// TwinCAT 3 PLC project BendingMachine
// ProgramVersion: 3.1.4026.27
// libraries:
//   Tc2_MC2, * (Beckhoff Automation GmbH)
//   Tc2_MC2_Drive, * (Beckhoff Automation GmbH)
//   Tc2_NCI, * (Beckhoff Automation GmbH)
//   Tc2_PlcInterpolation, * (Beckhoff Automation GmbH)
//   Tc2_Standard, * (Beckhoff Automation GmbH)
//   Tc2_SUPS, * (Beckhoff Automation GmbH)
//   Tc2_System, * (Beckhoff Automation GmbH)
//   Tc2_Utilities, * (Beckhoff Automation GmbH)
//   Tc3_JsonXml, * (Beckhoff Automation GmbH)
//   Tc3_MC2_AdvancedHoming, * (Beckhoff Automation GmbH)
// project tree:
//   DUTs/ ACTION_ENUM.TcDUT, AXIS_ENUM.TcDUT, CENTERING_ENUM.TcDUT, E_Alarm.TcDUT, EJECT_ENUM.TcDUT, OUTPUT_ACTION_ENUM.TcDUT, OUTPUT_ENUM.TcDUT, PRGSTATE_ENUM.TcDUT, ST_MpgEncoder.TcDUT, ST_TwoHandControl.TcDUT, TYPE_ACTION.TcDUT, TYPE_MACHINE_RX.TcDUT, TYPE_MACHINE_TX.TcDUT, TYPE_MACRO.TcDUT, TYPE_PARAMETERS.TcDUT, TYPE_POSITION.TcDUT, TYPE_SEQUENCE.TcDUT, TYPE_TASK.TcDUT
//   GVLs/ Alarms.TcGVL, Calibration.TcGVL, IO.TcGVL, Machine.TcGVL, ProgramDB.TcGVL, Safety.TcGVL, Size.TcGVL, Diag.TcGVL, Hmi.TcGVL
//   / PlcTask.TcTTO
//   POUs/ Clock.TcPOU, MAIN.TcPOU
//   Core/Valves/ SetMacro.TcPOU, WaitMacro.TcPOU, ST_Valve.TcDUT, ST_Input.TcDUT
//   POUs/Messages/ ClearAlarms.TcPOU, RaiseAlarm.TcPOU
//   POUs/MPG/ MPG_ReadStatus.TcPOU
//   Core/Nc/ FB_BuildGroups.TcPOU, FB_ClearInterpolationGroup.TcPOU, ST_AxisCfg.TcDUT, E_SeqCmd.TcDUT, E_SeqStep.TcDUT, FB_FeedTableBuilder.TcPOU, FB_SequenceRunner.TcPOU, E_NcChannelCmd.TcDUT, FB_NcChannels.TcPOU
//   POUs/TwoHand/ TwoHand_ReadStatus.TcPOU
//   Core/ Core_Param.TcGVL
//   Core/Cycle/ E_CycleState.TcDUT
//   Core/Diag/ E_CycleEndReason.TcDUT, ST_DiagEvent.TcDUT, ST_ChannelDiag.TcDUT, ST_Diag.TcDUT, FB_DiagLog.TcPOU
//   Core/Sync/ E_MFuncKind.TcDUT, E_MFuncOnError.TcDUT, ST_MFuncDef.TcDUT, F_MValve.TcPOU, F_MValveDirect.TcPOU, F_MSync.TcPOU, F_MSimple.TcPOU, FB_MFuncDispatcher.TcPOU
//   Machine/ E_Valve.TcDUT, Mach.TcGVL, FB_MachineConfig.TcPOU, FB_Centering.TcPOU, E_CenteringStep.TcDUT
//   Core/Axes/ FB_AxisModule.TcPOU, E_AxisAlarm.TcDUT
//   Core/Hmi/ E_HmiCommand.TcDUT, E_HmiResult.TcDUT, ST_HmiCmd.TcDUT, ST_HmiLive.TcDUT, ST_HmiAxisParam.TcDUT, ST_HmiParam.TcDUT, ST_HmiNamedItem.TcDUT, ST_HmiCfg.TcDUT, ST_HmiAxisSts.TcDUT, ST_HmiValveSts.TcDUT, ST_HmiSts.TcDUT, FB_HmiCommandHandler.TcPOU, FB_HmiWatchdog.TcPOU
// real-time tasks:
//   TASK PlcTask: cycle T#1ms, priority 20, ADS port 350
// motion (NC):
//   TASK NC-Task 1 SAF: cycle T#1ms, priority 1, ADS port 501
//   TASK NC-Task 1 SVB: cycle T#1ms, priority 8, ADS port 511
//   AXIS ERL (id 1)
//     General: UnitName=°
//     Dynamic: Acceleration=1780.713, Deceleration=1780.713, Jerk=5342.139
//     Velo: RefSearch=11.87142, RefSync=11.87142, SlowManual=59.3571, FastManual=356.1426, Fast=1187.142, Maximum=1187.142
//     OtherSettings: AllowMotionCmdToSlave=true
//     encoder EncType=8
//       EncPara: ScaleFactorNumerator=360, ScaleFactorDenominator=23068672, MaxCount=#xffffffff, ReferenceSystem=1
//         SoftEndMinControl: Enable=true, Range=-180
//         SoftEndMaxControl: Enable=true, Range=180
//     drive DrvType=9
//       DrvPara: MaxCount=#xffffffff, DriveControlDWord=#x00030100
//         Analog: VeloReferenz=1305.8562, VeloScale=1.02400649589962, TorqueSetpointScale=10, ScaleFactorActTorque=0.1
//         TimeComp: TaskDelayCycles=1
//     controller CtrType=1
//       CtrPara: PriorControlFactor=1
//         PosDiffControl: Enable=false
//         Observer: BandWidth=20
//   AXIS USEL (id 2)
//     Dynamic: Acceleration=1456.0155, Deceleration=1456.0155, Jerk=4368.0465
//     Velo: RefSearch=9.70677, RefSync=9.70677, SlowManual=12.5, FastManual=75, Fast=970.677, Maximum=970.677
//     OtherSettings: AllowMotionCmdToSlave=true
//     encoder EncType=8
//       EncPara: ScaleFactorNumerator=160, ScaleFactorDenominator=15728640, Offset=281.208719889323, Inverse=true, MaxCount=#xffffffff, ReferenceSystem=1
//         SoftEndMinControl: Enable=true, Range=66
//         SoftEndMaxControl: Enable=true, Range=1725
//     drive DrvType=9
//       DrvPara: Inverse=true, MaxCount=#xffffffff, DriveControlDWord=#x00030100
//         Analog: VeloReferenz=1067.7447, VeloScale=1.02400649589962, TorqueSetpointScale=10, ScaleFactorActTorque=0.1
//         TimeComp: TaskDelayCycles=1
//     controller CtrType=1
//       CtrPara: PriorControlFactor=1
//         Observer: BandWidth=20
//   AXIS ERR (id 3)
//     General: UnitName=°
//     Dynamic: Acceleration=1780.713, Deceleration=1780.713, Jerk=5342.139
//     Velo: RefSearch=11.87142, RefSync=11.87142, SlowManual=59.3571, FastManual=356.1426, Fast=1187.142, Maximum=1187.142
//     OtherSettings: AllowMotionCmdToSlave=true
//     encoder EncType=8
//       EncPara: ScaleFactorNumerator=360, ScaleFactorDenominator=23068672, Offset=78.9122668179599, MaxCount=#xffffffff, ReferenceSystem=1
//         SoftEndMinControl: Enable=true, Range=-180
//         SoftEndMaxControl: Enable=true, Range=180
//     drive DrvType=9
//       DrvPara: MaxCount=#xffffffff, DriveControlDWord=#x00030100
//         Analog: VeloReferenz=1305.8562, VeloScale=1.02400649589962, TorqueSetpointScale=10, ScaleFactorActTorque=0.1
//         TimeComp: TaskDelayCycles=1
//     controller CtrType=1
//       CtrPara: PriorControlFactor=1
//         Observer: BandWidth=20
//   AXIS USER (id 4)
//     Dynamic: Acceleration=1456.0155, Deceleration=1456.0155, Jerk=4368.0465
//     Velo: RefSearch=9.70677, RefSync=9.70677, SlowManual=12.5, FastManual=75, Fast=970.677, Maximum=970.677
//     OtherSettings: AllowMotionCmdToSlave=true
//     encoder EncType=8
//       EncPara: ScaleFactorNumerator=160, ScaleFactorDenominator=15728640, Offset=543.740122477214, Inverse=true, MaxCount=#xffffffff, ReferenceSystem=1
//         SoftEndMinControl: Enable=true, Range=66
//         SoftEndMaxControl: Enable=true, Range=1725
//     drive DrvType=9
//       DrvPara: Inverse=true, MaxCount=#xffffffff, DriveControlDWord=#x00030100
//         Analog: VeloReferenz=1067.7447, VeloScale=1.02400649589962, TorqueSetpointScale=10, ScaleFactorActTorque=0.1
//         TimeComp: TaskDelayCycles=1
//     controller CtrType=1
//       CtrPara: PriorControlFactor=1
//         Observer: BandWidth=20
//   AXIS UR (id 5)
//     General: UnitName=°
//     Dynamic: Acceleration=546.441, Deceleration=546.441, Jerk=1639.323
//     Velo: RefSearch=3.64294, RefSync=3.64294, SlowManual=18.2147, FastManual=109.2882, Fast=364.294, Maximum=364.294
//     OtherSettings: AllowMotionCmdToSlave=true
//     encoder EncType=8
//       EncPara: ScaleFactorNumerator=360, ScaleFactorDenominator=57671680, Offset=-105.826067837802, MaxCount=#xffffffff, ReferenceSystem=1
//         SoftEndMinControl: Enable=true, Range=-95
//         SoftEndMaxControl: Enable=true, Range=95
//     drive DrvType=9
//       DrvPara: MaxCount=#xffffffff, DriveControlDWord=#x00030100
//         Analog: VeloReferenz=400.7234, VeloScale=1.02400649589962, TorqueSetpointScale=10, ScaleFactorActTorque=0.1
//         TimeComp: TaskDelayCycles=1
//     controller CtrType=1
//       CtrPara: PriorControlFactor=1
//         Observer: BandWidth=20
//   AXIS UR SIM (id 6)
//     OtherSettings: AllowMotionCmdToSlave=true
//     encoder EncType=1
//     drive DrvType=5
//       Analog: TorqueSetpointScale=10, ScaleFactorActTorque=0.1
//       TimeComp: TaskDelayCycles=1
//     controller CtrType=1
//       CtrPara: PriorControlFactor=1
//         Observer: BandWidth=20
// I/O:
//   DEVICE Device 1 (EtherCAT), AmsNetId 192.168.1.106.2.1
//     Term 21 (EK1100) [EK1100 EtherCAT Coupler (2A E-Bus)]
//       Term 22 (EL6070-0033) [EL6070-0033 1Ch. Licence key terminal, individual licences]
//       Term 23 (EL1409) [EL1409 16Ch. Dig. Input 24V, 3ms]
//       Term 24 (EL1409) [EL1409 16Ch. Dig. Input 24V, 3ms]
//       Term 25 (EL2409) [EL2409 16Ch. Dig. Output 24V, 0.5A]
//       Term 26 (EK1322) [EK1322 2-port EtherCAT P junction with feed-in]
//         Box 27 (EPP1809-0022) [EPP1809-0022 16 Ch. Dig. Input 24V, 3ms, M8]
//         Box 28 (EPP1809-0022) [EPP1809-0022 16 Ch. Dig. Input 24V, 3ms, M8]
//       Term 29 (EL9410) [EL9410 E-Bus Power Supplier  (Diagnostics)]
//       Term 30 (EL6910) [EL6910, TwinSAFE PLC]
//       Term 31 (EL1918) [EL1918, 8Ch. Safety Input 24V, TwinSAFE]
//         modules: Module 1 (FSOE), Module 2 (FSLOGIC)
//       Term 32 (EL1918) [EL1918, 8Ch. Safety Input 24V, TwinSAFE]
//         modules: Module 1 (FSOE), Module 2 (FSLOGIC)
//       Term 33 (EL2904) [EL2904, 4 Ch. Safety Output 24V, 0.5A, TwinSAFE]
//         modules: Module 1 (FSOES), Module 2 (DO)
//       Term 34 (EK1110) [EK1110 EtherCAT extension]
//     Drive 35 (AX5206-0000-0216) [AX5206-0000-0216 EtherCAT Drive (SoE, 2 Ch.)]
//       Term 36 (AX5805) [AX5805 (Safety Drive Option)]
//         modules: Module 1 (Safety Process Data, 2 axis), Module 2 (Standard Process Data, 2 axis)
//     Drive 37 (AX5206-0000-0216) [AX5206-0000-0216 EtherCAT Drive (SoE, 2 Ch.)]
//       Term 38 (AX5805) [AX5805 (Safety Drive Option)]
//         modules: Module 1 (Safety Process Data, 2 axis), Module 2 (Standard Process Data, 2 axis)
//     Box 41 (EX260-SEC1) [EX260-SEC1 EtherCAT SI Unit (32DO_PNP) Rev1.2]
//     Box 42 (EX260-SEC1) [EX260-SEC1 EtherCAT SI Unit (32DO_PNP) Rev1.2]
//     Drive 39 (AX5103-0000-0216) [AX5103-0000-0216 EtherCAT Drive (SoE, 1 Ch.)]
//       Term 40 (AX5805) [AX5805 (Safety Drive Option)]
//         modules: Module 1 (Safety Process Data, 1 axis), Module 2 (Standard Process Data, 1 axis)
// variable links:
//   Device 1 (EtherCAT) <-> Device 1 (EtherCAT)/Drive 35 (AX5206-0000-0216)/Term 36 (AX5805)
//     Term 21 (EK1100)/Term 30 (EL6910)/ConnectionInputs/Message_184 TxPDO <-> Module 1 (Safety Process Data, 2 axis)/Outputs (Controlword)/FSOE
//     Term 21 (EK1100)/Term 30 (EL6910)/ConnectionOutputs/Message_184 RxPDO <-> Module 1 (Safety Process Data, 2 axis)/Inputs (Statusword)/FSOE
//   Device 1 (EtherCAT) <-> Device 1 (EtherCAT)/Drive 37 (AX5206-0000-0216)/Term 38 (AX5805)
//     Term 21 (EK1100)/Term 30 (EL6910)/ConnectionInputs/Message_183 TxPDO <-> Module 1 (Safety Process Data, 2 axis)/Outputs (Controlword)/FSOE
//     Term 21 (EK1100)/Term 30 (EL6910)/ConnectionOutputs/Message_183 RxPDO <-> Module 1 (Safety Process Data, 2 axis)/Inputs (Statusword)/FSOE
//   Device 1 (EtherCAT) <-> Device 1 (EtherCAT)/Drive 39 (AX5103-0000-0216)/Term 40 (AX5805)
//     Term 21 (EK1100)/Term 30 (EL6910)/ConnectionInputs/Message_191 TxPDO <-> Module 1 (Safety Process Data, 1 axis)/Outputs (Controlword)/FSOE
//     Term 21 (EK1100)/Term 30 (EL6910)/ConnectionOutputs/Message_191 RxPDO <-> Module 1 (Safety Process Data, 1 axis)/Inputs (Statusword)/FSOE
//   Device 1 (EtherCAT) <-> Device 1 (EtherCAT)/Term 21 (EK1100)/Term 31 (EL1918)
//     Term 21 (EK1100)/Term 30 (EL6910)/ConnectionInputs/Message_195 TxPDO <-> Module 1 (FSOE)/FSoE Outputs/FSOE
//     Term 21 (EK1100)/Term 30 (EL6910)/ConnectionOutputs/Message_195 RxPDO <-> Module 1 (FSOE)/FSoE Inputs/FSOE
//   Device 1 (EtherCAT) <-> Device 1 (EtherCAT)/Term 21 (EK1100)/Term 32 (EL1918)
//     Term 21 (EK1100)/Term 30 (EL6910)/ConnectionInputs/Message_196 TxPDO <-> Module 1 (FSOE)/FSoE Outputs/FSOE
//     Term 21 (EK1100)/Term 30 (EL6910)/ConnectionOutputs/Message_196 RxPDO <-> Module 1 (FSOE)/FSoE Inputs/FSOE
//   Device 1 (EtherCAT) <-> Device 1 (EtherCAT)/Term 21 (EK1100)/Term 33 (EL2904)
//     Term 21 (EK1100)/Term 30 (EL6910)/ConnectionInputs/Message_197 TxPDO <-> Module 1 (FSOES)/RxPDO/FSOE
//     Term 21 (EK1100)/Term 30 (EL6910)/ConnectionOutputs/Message_197 RxPDO <-> Module 1 (FSOES)/TxPDO/FSOE
//   NC-Task 1 SAF/Axes/ERL <-> Device 1 (EtherCAT)/Drive 35 (AX5206-0000-0216)
//     Drive/Inputs/In/nDataIn1 <-> AT 1/Following distance
//     Drive/Inputs/In/nDataIn3[0] <-> AT 1/Torque/force feedback value
//     Drive/Inputs/In/nDcOutputTime <-> InfoData/DcOutputShift
//     Drive/Inputs/In/nState1 <-> AT 1/Drive status word @bit 8
//     Drive/Inputs/In/nState2 <-> AT 1/Drive status word
//     Drive/Inputs/In/nState4 @bit 1 <-> WcState/InputToggle
//     Drive/Inputs/In/nState4 <-> WcState/WcState
//     Drive/Outputs/Out/nCtrl1 <-> MDT 1/Master control word @bit 8
//     Drive/Outputs/Out/nDataOut1 <-> MDT 1/Position command value
//     Enc/Inputs/In/nDataIn1 <-> AT 1/Position feedback 1 value
//     Enc/Inputs/In/nDcInputTime <-> InfoData/DcInputShift
//     Enc/Inputs/In/nState4 @bit 1 <-> WcState/InputToggle
//     Enc/Inputs/In/nState4 <-> WcState/WcState
//   NC-Task 1 SAF/Axes/ERR <-> Device 1 (EtherCAT)/Drive 37 (AX5206-0000-0216)
//     Drive/Inputs/In/nDataIn1 <-> AT 1/Following distance
//     Drive/Inputs/In/nDataIn3[0] <-> AT 1/Torque/force feedback value
//     Drive/Inputs/In/nDcOutputTime <-> InfoData/DcOutputShift
//     Drive/Inputs/In/nState1 <-> AT 1/Drive status word @bit 8
//     Drive/Inputs/In/nState2 <-> AT 1/Drive status word
//     Drive/Inputs/In/nState4 @bit 1 <-> WcState/InputToggle
//     Drive/Inputs/In/nState4 <-> WcState/WcState
//     Drive/Outputs/Out/nCtrl1 <-> MDT 1/Master control word @bit 8
//     Drive/Outputs/Out/nDataOut1 <-> MDT 1/Position command value
//     Enc/Inputs/In/nDataIn1 <-> AT 1/Position feedback 1 value
//     Enc/Inputs/In/nDcInputTime <-> InfoData/DcInputShift
//     Enc/Inputs/In/nState4 @bit 1 <-> WcState/InputToggle
//     Enc/Inputs/In/nState4 <-> WcState/WcState
//   NC-Task 1 SAF/Axes/UR <-> Device 1 (EtherCAT)/Drive 39 (AX5103-0000-0216)
//     Drive/Inputs/In/nDataIn1 <-> AT/Following distance
//     Drive/Inputs/In/nDataIn3[0] <-> AT/Torque/force feedback value
//     Drive/Inputs/In/nDcOutputTime <-> InfoData/DcOutputShift
//     Drive/Inputs/In/nState1 <-> AT/Drive status word @bit 8
//     Drive/Inputs/In/nState2 <-> AT/Drive status word
//     Drive/Inputs/In/nState4 @bit 1 <-> WcState/InputToggle
//     Drive/Inputs/In/nState4 <-> WcState/WcState
//     Drive/Outputs/Out/nCtrl1 <-> MDT/Master control word @bit 8
//     Drive/Outputs/Out/nDataOut1 <-> MDT/Position command value
//     Enc/Inputs/In/nDataIn1 <-> AT/Position feedback 1 value
//     Enc/Inputs/In/nDcInputTime <-> InfoData/DcInputShift
//     Enc/Inputs/In/nState4 @bit 1 <-> WcState/InputToggle
//     Enc/Inputs/In/nState4 <-> WcState/WcState
//   NC-Task 1 SAF/Axes/USEL <-> Device 1 (EtherCAT)/Drive 35 (AX5206-0000-0216)
//     Drive/Inputs/In/nDataIn1 <-> AT 2/Following distance
//     Drive/Inputs/In/nDataIn3[0] <-> AT 2/Torque/force feedback value
//     Drive/Inputs/In/nDcOutputTime <-> InfoData/DcOutputShift
//     Drive/Inputs/In/nState1 <-> AT 2/Drive status word @bit 8
//     Drive/Inputs/In/nState2 <-> AT 2/Drive status word
//     Drive/Inputs/In/nState4 @bit 1 <-> WcState/InputToggle
//     Drive/Inputs/In/nState4 <-> WcState/WcState
//     Drive/Outputs/Out/nCtrl1 <-> MDT 2/Master control word @bit 8
//     Drive/Outputs/Out/nDataOut1 <-> MDT 2/Position command value
//     Enc/Inputs/In/nDataIn1 <-> AT 2/Position feedback 1 value
//     Enc/Inputs/In/nDcInputTime <-> InfoData/DcInputShift
//     Enc/Inputs/In/nState4 @bit 1 <-> WcState/InputToggle
//     Enc/Inputs/In/nState4 <-> WcState/WcState
//   NC-Task 1 SAF/Axes/USER <-> Device 1 (EtherCAT)/Drive 37 (AX5206-0000-0216)
//     Drive/Inputs/In/nDataIn1 <-> AT 2/Following distance
//     Drive/Inputs/In/nDataIn3[0] <-> AT 2/Torque/force feedback value
//     Drive/Inputs/In/nDcOutputTime <-> InfoData/DcOutputShift
//     Drive/Inputs/In/nState1 <-> AT 2/Drive status word @bit 8
//     Drive/Inputs/In/nState2 <-> AT 2/Drive status word
//     Drive/Inputs/In/nState4 @bit 1 <-> WcState/InputToggle
//     Drive/Inputs/In/nState4 <-> WcState/WcState
//     Drive/Outputs/Out/nCtrl1 <-> MDT 2/Master control word @bit 8
//     Drive/Outputs/Out/nDataOut1 <-> MDT 2/Position command value
//     Enc/Inputs/In/nDataIn1 <-> AT 2/Position feedback 1 value
//     Enc/Inputs/In/nDcInputTime <-> InfoData/DcInputShift
//     Enc/Inputs/In/nState4 @bit 1 <-> WcState/InputToggle
//     Enc/Inputs/In/nState4 <-> WcState/WcState
//   BendingMachine/BendingMachine Instance <-> Device 1 (EtherCAT)/Box 41 (EX260-SEC1)
//     PlcTask Outputs/IO.smc1[{0..3}] <-> Byte {0..3}/Output  (4 links)
//   BendingMachine/BendingMachine Instance <-> Device 1 (EtherCAT)/Box 42 (EX260-SEC1)
//     PlcTask Outputs/IO.smc2[{0..3}] <-> Byte {0..3}/Output  (4 links)
//   BendingMachine/BendingMachine Instance <-> Device 1 (EtherCAT)/Drive 35 (AX5206-0000-0216)
//     PlcTask Inputs/MAIN.stMpgEncoder.diRowPositionFeedBack <-> AT 1/Position feedback 2 value (external feedback)
//   BendingMachine/BendingMachine Instance <-> Device 1 (EtherCAT)/Term 21 (EK1100)/Term 23 (EL1409)
//     PlcTask Inputs/IO.clampIn <-> DIP Inputs/Input Channel 14
//     PlcTask Inputs/IO.clampOpen <-> DIP Inputs/Input Channel 13
//     PlcTask Inputs/IO.fixedClampEncode <-> DIP Inputs/Input Channel 15
//     PlcTask Inputs/IO.mobileClampEncode <-> DIP Inputs/Input Channel 16
//     PlcTask Inputs/MAIN.stMpgEncoder.diButton1 <-> DIP Inputs/Input Channel 1
//     PlcTask Inputs/MAIN.stMpgEncoder.diButton2 <-> DIP Inputs/Input Channel 2
//     PlcTask Inputs/MAIN.stMpgEncoder.diButton3 <-> DIP Inputs/Input Channel 3
//     PlcTask Inputs/MAIN.stMpgEncoder.diSelector1Bit1 <-> DIP Inputs/Input Channel 4
//     PlcTask Inputs/MAIN.stMpgEncoder.diSelector1Bit2 <-> DIP Inputs/Input Channel 5
//     PlcTask Inputs/MAIN.stMpgEncoder.diSelector1Bit3 <-> DIP Inputs/Input Channel 6
//     PlcTask Inputs/MAIN.stMpgEncoder.diSelector2Bit1 <-> DIP Inputs/Input Channel 7
//     PlcTask Inputs/MAIN.stMpgEncoder.diSelector2Bit2 <-> DIP Inputs/Input Channel 8
//     PlcTask Inputs/MAIN.stTwoHandControl.diStartButton <-> DIP Inputs/Input Channel 9
//     PlcTask Inputs/MAIN.stTwoHandControl.diStopButton <-> DIP Inputs/Input Channel 10
//     PlcTask Inputs/Safety.PulsanteResetBarriere <-> DIP Inputs/Input Channel 12
//     PlcTask Inputs/Safety.PulsanteResetEmergenza <-> DIP Inputs/Input Channel 11
//   BendingMachine/BendingMachine Instance <-> Device 1 (EtherCAT)/Term 21 (EK1100)/Term 24 (EL1409)
//     PlcTask Inputs/IO.cabinetThermostat <-> DIP Inputs/Input Channel 10
//     PlcTask Inputs/IO.chillerAlarm <-> DIP Inputs/Input Channel 5
//     PlcTask Inputs/IO.chillerMagnetTrip <-> DIP Inputs/Input Channel 6
//     PlcTask Inputs/IO.doorLeftClosed <-> DIP Inputs/Input Channel 7
//     PlcTask Inputs/IO.doorRightClosed <-> DIP Inputs/Input Channel 8
//     PlcTask Inputs/IO.fuseAlarm <-> DIP Inputs/Input Channel 1
//     PlcTask Inputs/IO.leftAxisMagnetTrip <-> DIP Inputs/Input Channel 2
//     PlcTask Inputs/IO.pressureSwMinPressure <-> DIP Inputs/Input Channel 9
//     PlcTask Inputs/IO.rightAxisMagnetTrip <-> DIP Inputs/Input Channel 3
//     PlcTask Inputs/IO.ur2MagnetTrip <-> DIP Inputs/Input Channel 4
//   BendingMachine/BendingMachine Instance <-> Device 1 (EtherCAT)/Term 21 (EK1100)/Term 25 (EL2409)
//     PlcTask Outputs/IO.chillerEnabled <-> Channel 10/Output
//     PlcTask Outputs/IO.fuseReset <-> Channel 9/Output
//     PlcTask Outputs/IO.spiaPulsanteStart <-> Channel 7/Output
//     PlcTask Outputs/IO.spiaPulsanteStop <-> Channel 8/Output
//     PlcTask Outputs/IO.turretGreen <-> Channel 2/Output
//     PlcTask Outputs/IO.turretRed <-> Channel 1/Output
//     PlcTask Outputs/IO.turretSiren <-> Channel 4/Output
//     PlcTask Outputs/IO.turretYellow <-> Channel 3/Output
//     PlcTask Outputs/Safety.SpiaPulsanteRipristinoBarriere <-> Channel 6/Output
//     PlcTask Outputs/Safety.SpiaPulsanteRipristinoSicurezze <-> Channel 5/Output
//   BendingMachine/BendingMachine Instance <-> Device 1 (EtherCAT)/Term 21 (EK1100)/Term 26 (EK1322)/Box 27 (EPP1809-0022)
//     PlcTask Inputs/IO.centering1LeftIn <-> Channel 10/Input
//     PlcTask Inputs/IO.centering2LeftIn <-> Channel 9/Input
//     PlcTask Inputs/IO.centering3LeftIn <-> Channel 12/Input
//     PlcTask Inputs/IO.centering4LeftIn <-> Channel 11/Input
//     PlcTask Inputs/IO.epLeftBendUp <-> Channel 6/Input
//     PlcTask Inputs/IO.epLeftIn <-> Channel 5/Input
//     PlcTask Inputs/IO.erLeftIn <-> Channel 4/Input
//     PlcTask Inputs/IO.erLeftOut <-> Channel 3/Input
//     PlcTask Inputs/IO.useLeftDown <-> Channel 2/Input
//     PlcTask Inputs/IO.useLeftUp <-> Channel 1/Input
//   BendingMachine/BendingMachine Instance <-> Device 1 (EtherCAT)/Term 21 (EK1100)/Term 26 (EK1322)/Box 28 (EPP1809-0022)
//     PlcTask Inputs/IO.epRightBendUp <-> Channel 6/Input
//     PlcTask Inputs/IO.epRightIn <-> Channel 5/Input
//     PlcTask Inputs/IO.erRightIn <-> Channel 4/Input
//     PlcTask Inputs/IO.erRightOut <-> Channel 3/Input
//     PlcTask Inputs/IO.useRightDown <-> Channel 2/Input
//     PlcTask Inputs/IO.useRighttUp <-> Channel 1/Input
//   BendingMachine/BendingMachine Instance <-> Device 1 (EtherCAT)/Term 21 (EK1100)/Term 30 (EL6910)
//     PlcTask Inputs/MAIN.stMpgEncoder.diSafetySwitch <-> StandardInputs/Standard Out Var 64
//     PlcTask Inputs/MAIN.stTwoHandControl.diSafetySwitch <-> StandardInputs/Standard Out Var 60
//     PlcTask Inputs/MAIN.stTwoHandControl.diTwoHand <-> StandardInputs/Standard Out Var 65
//     PlcTask Inputs/Safety.AbilitazionePeriferiche <-> StandardInputs/Standard Out Var 50
//     PlcTask Inputs/Safety.BarriereResettate <-> StandardInputs/Standard Out Var 62
//     PlcTask Inputs/Safety.ComErr <-> StandardInputs/Standard Out Var 13
//     PlcTask Inputs/Safety.ComStartup <-> StandardInputs/Standard Out Var 14
//     PlcTask Inputs/Safety.ERL_Error <-> StandardInputs/Standard Out Var 93
//     PlcTask Inputs/Safety.ERL_SDI_n <-> StandardInputs/Standard Out Var 92
//     PlcTask Inputs/Safety.ERL_SDI_p <-> StandardInputs/Standard Out Var 91
//     PlcTask Inputs/Safety.ERL_SOS <-> StandardInputs/Standard Out Var 89
//     PlcTask Inputs/Safety.ERL_SSM1 <-> StandardInputs/Standard Out Var 87
//     PlcTask Inputs/Safety.ERL_SSM2 <-> StandardInputs/Standard Out Var 88
//     PlcTask Inputs/Safety.ERL_SSR <-> StandardInputs/Standard Out Var 90
//     PlcTask Inputs/Safety.ERL_STO <-> StandardInputs/Standard Out Var 86
//     PlcTask Inputs/Safety.ERR_Error <-> StandardInputs/Standard Out Var 112
//     PlcTask Inputs/Safety.ERR_SDI_n <-> StandardInputs/Standard Out Var 113
//     PlcTask Inputs/Safety.ERR_SDI_p <-> StandardInputs/Standard Out Var 103
//     PlcTask Inputs/Safety.ERR_SOS <-> StandardInputs/Standard Out Var 104
//     PlcTask Inputs/Safety.ERR_SSM1 <-> StandardInputs/Standard Out Var 105
//     PlcTask Inputs/Safety.ERR_SSM2 <-> StandardInputs/Standard Out Var 106
//     PlcTask Inputs/Safety.ERR_SSR <-> StandardInputs/Standard Out Var 107
//     PlcTask Inputs/Safety.ERR_SSR2 <-> StandardInputs/Standard Out Var 182
//     PlcTask Inputs/Safety.ERR_STO <-> StandardInputs/Standard Out Var 108
//     PlcTask Inputs/Safety.EmergenzaResettata <-> StandardInputs/Standard Out Var 19
//     PlcTask Inputs/Safety.FBDeactivate <-> StandardInputs/Standard Out Var 15
//     PlcTask Inputs/Safety.FBErr <-> StandardInputs/Standard Out Var 12
//     PlcTask Inputs/Safety.FBRun <-> StandardInputs/Standard Out Var 16
//     PlcTask Inputs/Safety.InRun <-> StandardInputs/Standard Out Var 18
//     PlcTask Inputs/Safety.ModoAuto1Op <-> StandardInputs/Standard Out Var 45
//     PlcTask Inputs/Safety.ModoAuto2Op <-> StandardInputs/Standard Out Var 163
//     PlcTask Inputs/Safety.ModoManuale <-> StandardInputs/Standard Out Var 46
//     PlcTask Inputs/Safety.ModoSemiAuto <-> StandardInputs/Standard Out Var 61
//     PlcTask Inputs/Safety.OtherErr <-> StandardInputs/Standard Out Var 17
//     PlcTask Inputs/Safety.SSR1_Enable <-> StandardInputs/Standard Out Var 179
//     PlcTask Inputs/Safety.SSR2_Enable <-> StandardInputs/Standard Out Var 180
//     PlcTask Inputs/Safety.UR_ComErr <-> StandardInputs/Standard Out Var 144
//     PlcTask Inputs/Safety.UR_ComStartup <-> StandardInputs/Standard Out Var 145
//     PlcTask Inputs/Safety.UR_Error <-> StandardInputs/Standard Out Var 136
//     PlcTask Inputs/Safety.UR_FBDeactivate <-> StandardInputs/Standard Out Var 146
//     PlcTask Inputs/Safety.UR_FBErr <-> StandardInputs/Standard Out Var 147
//     PlcTask Inputs/Safety.UR_FBRun <-> StandardInputs/Standard Out Var 149
//     PlcTask Inputs/Safety.UR_InRun <-> StandardInputs/Standard Out Var 148
//     PlcTask Inputs/Safety.UR_OtherErr <-> StandardInputs/Standard Out Var 150
//     PlcTask Inputs/Safety.UR_SDI_n <-> StandardInputs/Standard Out Var 137
//     PlcTask Inputs/Safety.UR_SDI_p <-> StandardInputs/Standard Out Var 138
//     PlcTask Inputs/Safety.UR_SOS <-> StandardInputs/Standard Out Var 139
//     PlcTask Inputs/Safety.UR_SSM1 <-> StandardInputs/Standard Out Var 140
//     PlcTask Inputs/Safety.UR_SSM2 <-> StandardInputs/Standard Out Var 141
//     PlcTask Inputs/Safety.UR_SSR <-> StandardInputs/Standard Out Var 142
//     PlcTask Inputs/Safety.UR_STO <-> StandardInputs/Standard Out Var 143
//     PlcTask Inputs/Safety.USEL_ERL_ComErr <-> StandardInputs/Standard Out Var 95
//     PlcTask Inputs/Safety.USEL_ERL_ComStartup <-> StandardInputs/Standard Out Var 96
//     PlcTask Inputs/Safety.USEL_ERL_FBDeactivate <-> StandardInputs/Standard Out Var 97
//     PlcTask Inputs/Safety.USEL_ERL_FBErr <-> StandardInputs/Standard Out Var 98
//     PlcTask Inputs/Safety.USEL_ERL_FBRun <-> StandardInputs/Standard Out Var 100
//     PlcTask Inputs/Safety.USEL_ERL_InRun <-> StandardInputs/Standard Out Var 99
//     PlcTask Inputs/Safety.USEL_ERL_OtherErr <-> StandardInputs/Standard Out Var 101
//     PlcTask Inputs/Safety.USEL_Error <-> StandardInputs/Standard Out Var 117
//     PlcTask Inputs/Safety.USEL_SDI_n <-> StandardInputs/Standard Out Var 118
//     PlcTask Inputs/Safety.USEL_SDI_p <-> StandardInputs/Standard Out Var 119
//     PlcTask Inputs/Safety.USEL_SOS <-> StandardInputs/Standard Out Var 120
//     PlcTask Inputs/Safety.USEL_SSM1 <-> StandardInputs/Standard Out Var 121
//     PlcTask Inputs/Safety.USEL_SSM2 <-> StandardInputs/Standard Out Var 122
//     PlcTask Inputs/Safety.USEL_SSR <-> StandardInputs/Standard Out Var 123
//     PlcTask Inputs/Safety.USEL_STO <-> StandardInputs/Standard Out Var 124
//     PlcTask Inputs/Safety.USER_ERR_ComErr <-> StandardInputs/Standard Out Var 102
//     PlcTask Inputs/Safety.USER_ERR_ComStartup <-> StandardInputs/Standard Out Var 111
//     PlcTask Inputs/Safety.USER_ERR_FBDeactivate <-> StandardInputs/Standard Out Var 109
//     PlcTask Inputs/Safety.USER_ERR_FBErr <-> StandardInputs/Standard Out Var 110
//     PlcTask Inputs/Safety.USER_ERR_FBRun <-> StandardInputs/Standard Out Var 115
//     PlcTask Inputs/Safety.USER_ERR_InRun <-> StandardInputs/Standard Out Var 114
//     PlcTask Inputs/Safety.USER_ERR_OtherErr <-> StandardInputs/Standard Out Var 116
//     PlcTask Inputs/Safety.USER_Error <-> StandardInputs/Standard Out Var 125
//     PlcTask Inputs/Safety.USER_SDI_n <-> StandardInputs/Standard Out Var 126
//     PlcTask Inputs/Safety.USER_SDI_p <-> StandardInputs/Standard Out Var 135
//     PlcTask Inputs/Safety.USER_SOS <-> StandardInputs/Standard Out Var 127
//     PlcTask Inputs/Safety.USER_SSM1 <-> StandardInputs/Standard Out Var 128
//     PlcTask Inputs/Safety.USER_SSM2 <-> StandardInputs/Standard Out Var 129
//     PlcTask Inputs/Safety.USER_SSR <-> StandardInputs/Standard Out Var 130
//     PlcTask Inputs/Safety.USER_SSR2 <-> StandardInputs/Standard Out Var 181
//     PlcTask Inputs/Safety.USER_STO <-> StandardInputs/Standard Out Var 131
//     PlcTask Outputs/Safety.Ack <-> StandardOutputs/Standard In Var 1
//     PlcTask Outputs/Safety.ModuleFault <-> StandardOutputs/Standard In Var 58
//     PlcTask Outputs/Safety.ResetBarriere <-> StandardOutputs/Standard In Var 63
//     PlcTask Outputs/Safety.ResetEmergenza <-> StandardOutputs/Standard In Var 31
//     PlcTask Outputs/Safety.Run <-> StandardOutputs/Standard In Var 2
//     PlcTask Outputs/Safety.UR_Ack <-> StandardOutputs/Standard In Var 81
//     PlcTask Outputs/Safety.UR_Run <-> StandardOutputs/Standard In Var 82
//     PlcTask Outputs/Safety.USEL_ERL_Ack <-> StandardOutputs/Standard In Var 76
//     PlcTask Outputs/Safety.USEL_ERL_Run <-> StandardOutputs/Standard In Var 77
//     PlcTask Outputs/Safety.USER_ERR_Ack <-> StandardOutputs/Standard In Var 79
//     PlcTask Outputs/Safety.USER_ERR_Run <-> StandardOutputs/Standard In Var 80
//   BendingMachine/BendingMachine Instance <-> NC-Task 1 SAF/Axes/ERL
//     PlcTask Inputs/MAIN.ERL.NcToPlc <-> Outputs/ToPlc
//     PlcTask Outputs/MAIN.ERL.PlcToNc <-> Inputs/FromPlc
//   BendingMachine/BendingMachine Instance <-> NC-Task 1 SAF/Axes/ERR
//     PlcTask Inputs/MAIN.ERR.NcToPlc <-> Outputs/ToPlc
//     PlcTask Outputs/MAIN.ERR.PlcToNc <-> Inputs/FromPlc
//   BendingMachine/BendingMachine Instance <-> NC-Task 1 SAF/Axes/UR
//     PlcTask Inputs/MAIN.UR2.NcToPlc <-> Outputs/ToPlc
//     PlcTask Outputs/MAIN.UR2.PlcToNc <-> Inputs/FromPlc
//   BendingMachine/BendingMachine Instance <-> NC-Task 1 SAF/Axes/UR SIM
//     PlcTask Inputs/MAIN.UR_SIM.NcToPlc <-> Outputs/ToPlc
//     PlcTask Outputs/MAIN.UR_SIM.PlcToNc <-> Inputs/FromPlc
//   BendingMachine/BendingMachine Instance <-> NC-Task 1 SAF/Axes/USEL
//     PlcTask Inputs/MAIN.USEL.NcToPlc <-> Outputs/ToPlc
//     PlcTask Outputs/MAIN.USEL.PlcToNc <-> Inputs/FromPlc
//   BendingMachine/BendingMachine Instance <-> NC-Task 1 SAF/Axes/USER
//     PlcTask Inputs/MAIN.USER.NcToPlc <-> Outputs/ToPlc
//     PlcTask Outputs/MAIN.USER.PlcToNc <-> Inputs/FromPlc
//   BendingMachine/BendingMachine Instance <-> NC-Task 1 SAF/Channel 1
//     PlcTask Inputs/MAIN.in_stNciToPlc[0] <-> Outputs/ToPlc
//     PlcTask Outputs/MAIN.out_stPlcToNci[0] <-> Inputs/FromPlc
//   BendingMachine/BendingMachine Instance <-> NC-Task 1 SAF/Channel 2
//     PlcTask Inputs/MAIN.in_stNciToPlc[1] <-> Outputs/ToPlc
//     PlcTask Outputs/MAIN.out_stPlcToNci[1] <-> Inputs/FromPlc
//   BendingMachine/BendingMachine Instance <-> NC-Task 1 SAF/Channel 3
//     PlcTask Inputs/MAIN.in_stNciToPlc[2] <-> Outputs/ToPlc
//     PlcTask Outputs/MAIN.out_stPlcToNci[2] <-> Inputs/FromPlc

CONFIGURATION BendingMachine
    RESOURCE PLC ON TwinCAT3
        TASK PlcTask(INTERVAL := T#1ms, PRIORITY := 20);
        PROGRAM MAIN WITH PlcTask : MAIN;
    END_RESOURCE
END_CONFIGURATION

// ---- DUTs/ACTION_ENUM.TcDUT
{attribute 'qualified_only'}
{attribute 'strict'}
TYPE ACTION_ENUM :
(
	null 		:= 0,
	MOVEMENT 	:= 1,
	MACRO 		:= 2
);
END_TYPE

// ---- DUTs/AXIS_ENUM.TcDUT
{attribute 'qualified_only'}
{attribute 'strict'}
TYPE AXIS_ENUM :
(
	null := 0,
	USEL := 1,
	USER := 2,
	ERL := 3,
	ERR := 4,
	UR2 := 5,
	UR_SIM := 6
)UDINT;
END_TYPE

// ---- DUTs/CENTERING_ENUM.TcDUT
{attribute 'qualified_only'}
{attribute 'strict'}
TYPE CENTERING_ENUM :
(
	NO 	:= 0,
	TL	:= 1,
	TB	:= 2,
	ACC := 3
);
END_TYPE

// ---- DUTs/E_Alarm.TcDUT
// Indice degli allarmi in Alarms.Active / Alarms.Info.
// I testi (titolo, causa, rimedio) sono nell'HMI: chiavi Ui.Alarm.<numero>.*
// Un numero non si riusa mai per un significato diverso: l'HMI e lo storico allarmi lo usano come codice.
// Niente 'strict': i valori servono da indice di array.
{attribute 'qualified_only'}
TYPE E_Alarm :
(
	// --- Sicurezza (a livello) ---
	EmergencyStop := 1,	// circuito di emergenza non ripristinato
	DoorLeftOpen := 2,	// portiera sinistra aperta
	DoorRightOpen := 3,	// portiera destra aperta
	LightCurtainNotReset := 4,	// barriere fotoelettriche da ripristinare
	SafetyMainGroupError := 5,	// errore gruppo TwinSAFE principale
	SafetyGroupLeftError := 6,	// errore gruppo TwinSAFE USE SX / ER SX
	SafetyGroupRightError := 7,	// errore gruppo TwinSAFE USE DX / ER DX
	SafetyGroupUrError := 8,	// errore gruppo TwinSAFE UR
	// --- Azionamenti (a livello, Info = ErrorCode NC) ---
	DriveErl := 20,	// azionamento ER SX in errore
	DriveUsel := 21,	// azionamento USE SX in errore
	DriveUr2 := 22,	// azionamento UR2 in errore
	DriveErr := 23,	// azionamento ER DX in errore
	DriveUser := 24,	// azionamento USE DX in errore
	// --- Quadro elettrico (a livello, ingresso TRUE = guasto, bloccano lo start) ---
	FuseTripped := 40,	// fusibile intervenuto
	BreakerLeftAxis := 41,	// magnetotermico assi lato sinistro
	BreakerRightAxis := 42,	// magnetotermico assi lato destro
	BreakerUr2 := 43,	// magnetotermico UR2
	BreakerChiller := 44,	// magnetotermico climatizzatore
	AirPressureLow := 45,	// pressione aria sotto il minimo
	// --- Ciclo (memorizzati fino al Reset) ---
	CycleResetRequired := 60,	// ciclo interrotto: eseguire il Reset
	CenteringPartAlreadyPresent := 61,	// centratore: pezzo gia' presente prima della ricerca (passo 62)
	CenteringPartNotFound := 62,	// centratore: pezzo non trovato entro la corsa massima (passo 65)
	StartDriveError := 63,	// start rifiutato: azionamento in errore
	StartMotorsOff := 64,	// start rifiutato: motori non attivi
	StartNoProgram := 65,	// start rifiutato: nessun programma caricato
	StartCabinetAlarm := 66,	// start rifiutato: allarme quadro elettrico
	CenteringModeNotSupported := 67,	// modo di centraggio non gestito dal PLC (es. ACC); Info = valore di centering (passo 50)
	UnknownMFunction := 68,	// funzione M non gestita: il canale resterebbe fermo; Info = canale*1000 + M (1 SX, 2 DX, 3 UR2)
	StateTimeout := 69,	// passo tecnico del ciclo (reset/costruzione gruppi, tabelle, stop, reset assi) bloccato; Info = passo
	// --- Avvisi (non bloccanti) ---
	BatchCompleted := 90,	// lotto completato (contapezzi raggiunto)
	ChillerAlarm := 91,	// climatizzatore quadro in allarme
	CabinetOverTemperature := 92,	// temperatura quadro elevata
	// --- Timeout movimenti (Info = numero funzione M) ---
	ErLeftUp := 100,	// ER SX salita (M40)
	ErLeftDown := 101,	// ER SX discesa (M41)
	ErRightUp := 102,	// ER DX salita (M42)
	ErRightDown := 103,	// ER DX discesa (M43)
	UseLeftUp := 104,	// USE SX salita (M44)
	UseLeftDown := 105,	// USE SX discesa (M45)
	UseRightUp := 106,	// USE DX salita (M46)
	UseRightDown := 107,	// USE DX discesa (M47)
	SupportLeftOut := 108,	// spallamento SX uscita (M50)
	SupportLeftIn := 109,	// spallamento SX rientro (M51)
	SupportRightOut := 110,	// spallamento DX uscita (M48)
	SupportRightIn := 111,	// spallamento DX rientro (M49)
	EpLeftBend := 112,	// EP SX trazione (M70)
	EpLeftOut := 113,	// EP SX uscita (M72)
	EpLeftIn := 114,	// EP SX rientro (M73)
	EpLeftBendReturn := 115,	// EP SX ritorno trazione (M74)
	EpRightBend := 116,	// EP DX trazione (M70)
	EpRightOut := 117,	// EP DX uscita (M72)
	EpRightIn := 118,	// EP DX rientro (M73)
	EpRightBendReturn := 119,	// EP DX ritorno trazione (M74)
	// Attese di sincronismo e di espulsione: 15 s con il ciclo fermo su quell'attesa (MacroManager)
	SyncLeftWaitRight := 120,	// USE SX aspetta la USE DX (M61)
	SyncRightWaitLeft := 121,	// USE DX aspetta la USE SX (M60)
	SyncLeftWaitUr2 := 122,	// USE SX aspetta l'UR2 (M80)
	SyncRightWaitUr2 := 123,	// USE DX aspetta l'UR2 (M80)
	SyncLeftWaitUr2Ack := 124,	// USE SX aspetta che l'UR2 riceva la conferma (M112)
	SyncRightWaitUr2Ack := 125,	// USE DX aspetta che l'UR2 riceva la conferma (M113)
	SyncUr2WaitUseAck := 126,	// UR2 aspetta la conferma delle due USE (M110)
	SyncUr2WaitUse := 127,	// UR2 aspetta il posizionamento delle due USE (M116)
	EjectUr2NotAtZero := 128,	// espulsione: UR2 non a zero (M102)
	// --- Calibrazione e scrittura parametri (Info = ErrorID) ---
	HomingErl := 160,	// calibrazione ER SX fallita
	HomingUsel := 161,	// calibrazione USE SX fallita
	HomingUr2 := 162,	// calibrazione UR2 fallita
	HomingErr := 163,	// calibrazione ER DX fallita
	HomingUser := 164,	// calibrazione USE DX fallita
	ParamWriteErl := 170,	// scrittura limiti ER SX fallita
	ParamWriteUsel := 171,	// scrittura limiti USE SX fallita
	ParamWriteUr2 := 172,	// scrittura limiti UR2 fallita
	ParamWriteErr := 173,	// scrittura limiti ER DX fallita
	ParamWriteUser := 174,	// scrittura limiti USE DX fallita
	// --- Errori NC interni (Info = ErrorID NC) ---
	NcCenteringClearGroup := 200,	// centratore: reset gruppi (passo 55)
	NcCenteringApproach := 201,	// centratore: avvicinamento (passo 61)
	NcCenteringSearch := 202,	// centratore: ricerca pezzo (passo 65)
	NcCenteringStopSearch := 203,	// centratore: arresto dopo pezzo trovato (passo 67)
	NcCenteringStop := 204,	// centratore: arresto finale (passo 72)
	NcCenteringExtra := 205,	// centratore: posizionamento extra (passo 76)
	NcClearGroups := 206,	// reset gruppi di interpolazione (passo 120)
	NcClearGroupsInit := 207,	// reset gruppi di interpolazione INIT (passo 122)
	NcBuildGroups := 208,	// costruzione gruppi (passo 120)
	NcBuildGroupsInit := 209,	// costruzione gruppi INIT (passo 122)
	NcFeedTableReset := 210,	// reset tabelle avanzamento (passo 120)
	NcFeedTableResetInit := 211,	// reset tabelle avanzamento INIT (passo 122)
	NcFeedTablePrep := 212,	// preparazione tabelle avanzamento (passo 120)
	NcFeedTablePrepInit := 213,	// preparazione tabelle avanzamento INIT (passo 122)
	NcFeedTableStart := 214,	// avvio tabelle avanzamento (passo 120)
	NcFeedTableStartInit := 215,	// avvio tabelle avanzamento INIT (passo 122)
	NcFeedTableRun := 216,	// tabella avanzamento durante il ciclo (passo 410)
	NcFeedTableRunInit := 217,	// tabella avanzamento durante INIT (passo 412)
	NcAbort := 218,	// arresto di emergenza NC in abort (passo 600)
	NcStop := 219,	// arresto NC in stop (passo 700)
	NcStepOn := 220,	// ripartenza dopo stop (passo 730)
	NcResetAxes := 221,	// reset assi (passo 800)
	NcManualEStop := 222,	// passaggio in manuale: arresto NC (passo 905)
	NcManualClearGroup := 223,	// passaggio in manuale: reset gruppi (passo 910)
	NcManualResetAxes := 224,	// passaggio in manuale: reset assi (passo 920)
	NcResumeReset := 225	// ripresa dopo stop fuori dal RUN: reset canali NC (passo 745)
) UINT;
END_TYPE

// ---- DUTs/EJECT_ENUM.TcDUT
{attribute 'qualified_only'}
{attribute 'strict'}
TYPE EJECT_ENUM :
(
	YES := 0,
	NO_2_START := 1,
	NO_1_START := 2
)UDINT;
END_TYPE

// ---- DUTs/OUTPUT_ACTION_ENUM.TcDUT
{attribute 'qualified_only'}
{attribute 'strict'}
TYPE OUTPUT_ACTION_ENUM :
(
	SET := 0,
	RESET := 1
);
END_TYPE

// ---- DUTs/OUTPUT_ENUM.TcDUT
{attribute 'qualified_only'}
{attribute 'strict'}
TYPE OUTPUT_ENUM :
(
	MONOSTABLE := 0,
	BISTABLE := 1
);
END_TYPE

// ---- DUTs/PRGSTATE_ENUM.TcDUT
{attribute 'qualified_only'}
{attribute 'strict'}
TYPE PRGSTATE_ENUM :
(
	FREE := 0,
	RESET := 1,
	ACTIVE := 2,
	END := 3,
	STOP := 4
);
END_TYPE

// ---- DUTs/ST_MpgEncoder.TcDUT
TYPE ST_MpgEncoder :
STRUCT
	diButton1				 AT %I* : BOOL;
	diButton2				 AT %I* : BOOL;
	diButton3				 AT %I* : BOOL;
	diSelector1Bit1			 AT %I* : BOOL;
	diSelector1Bit2			 AT %I* : BOOL;
	diSelector1Bit3			 AT %I* : BOOL;
	diSelector2Bit1		     AT %I* : BOOL;
	diSelector2Bit2		     AT %I* : BOOL;
	diSafetySwitch		     AT %I* : BOOL;
	diSelector1						: BYTE;
	diSelector2						: BYTE;
	diRowPositionFeedBack	 AT %I* : DINT;
	rActPos							: REAL;
	rActVelo						: REAL;
	uiOverrideSpeed					: UINT;
	eDirection						: MC_Direction;
	tUpdateTime						: TIME;
	uiScalingFactorNumerator		: UINT;
	uiScalingFactorDenominator		: UINT;
	uiSpeedDivider					: UINT;
	uiMaxSpeed						: UINT := 5;
	xButton1RTrigger				: BOOL;
	xButton2RTrigger				: BOOL;
	xButton3RTrigger				: BOOL;
	xFowardRTrigger					: BOOL;
	xBackwardRTrigger				: BOOL;
	xSafetySwitchRTrigger			: BOOL;
	xButton1FTrigger				: BOOL;
	xButton2FTrigger				: BOOL;
	xButton3FTrigger				: BOOL;
	xFowardFTrigger					: BOOL;
	xBackwardFTrigger				: BOOL;
	xSafetySwitchFTrigger			: BOOL;
END_STRUCT
END_TYPE

// ---- DUTs/ST_TwoHandControl.TcDUT
TYPE ST_TwoHandControl :
STRUCT
	diButton1		 AT %I* : BOOL;
	diStartButton	 AT %I* : BOOL;
	diStopButton	 AT %I* : BOOL;
	diTwoHand		 AT %I* : BOOL;
	diTwoHand1		 AT %I* : BOOL;
	diTwoHand2		 AT %I* : BOOL;
	diSafetySwitch	 AT %I* : BOOL;
	doStartLED		 AT %Q* : BOOL;
	doStopLED		 AT %Q* : BOOL;
	
	xButton1RTrigger		: BOOL;
	xButton1FTrigger		: BOOL;
	xStartRTrigger			: BOOL;
	xStartFTrigger			: BOOL;
	xStopRTrigger			: BOOL;
	xStopFTrigger			: BOOL;
	xTwoHandRTrigger		: BOOL;
	xTwoHandFTRigger		: BOOL;
	xSafetySwitchRTrigger	: BOOL;
	xSafetySwitchFTrigger	: BOOL;
	xStopButtonDelayTrigger	: BOOL;
END_STRUCT
END_TYPE

// ---- DUTs/TYPE_ACTION.TcDUT
TYPE TYPE_ACTION :
STRUCT
	active : BOOL;
	speed : UDINT;
	lineNo : UDINT;
	aType : ACTION_ENUM;
	centeringVerse : DINT;
	centeringAmount : LREAL;
	autoCorrection : BOOL;
	pos : ARRAY[0..Size.MAX_POSITION-1] OF TYPE_POSITION;
	macros : ARRAY[0..Size.MAX_MACRO-1] OF TYPE_MACRO;
END_STRUCT
END_TYPE

// ---- DUTs/TYPE_MACHINE_RX.TcDUT
TYPE TYPE_MACHINE_RX :
STRUCT
	ERLCalibrated			: BOOL;
	USELCalibrated			: BOOL;
	UR2Calibrated			: BOOL;
	ERRCalibrated			: BOOL;
	USERCalibrated			: BOOL;
	ERLPresent				: BOOL;
	USELPresent				: BOOL;
	UR2Present				: BOOL;
	ERRPresent				: BOOL;
	USERPresent				: BOOL;
	ERLCheckDone			: BOOL;
	USELCheckDone			: BOOL;
	ER2CheckDone			: BOOL;
	ERRCheckDone			: BOOL;
	USERCheckDone			: BOOL;
	EnableSirenOverride		: BOOL;
	UseLUpperLimit			: LREAL;
	UseLLowerLimit			: LREAL;
	UseRUpperLimit			: LREAL;
	UseRLowerLimit			: LREAL;
	ErLUpperLimit			: LREAL;
	ErLLowerLimit			: LREAL;
	ErRUpperLimit			: LREAL;
	ErRLowerLimit			: LREAL;
	UrRUpperLimit			: LREAL;
	UrRLowerLimit			: LREAL;
END_STRUCT
END_TYPE

// ---- DUTs/TYPE_MACHINE_TX.TcDUT
TYPE TYPE_MACHINE_TX :
STRUCT
	lastERLKnownPosition	: LREAL;
	lastUSELKnownPosition	: LREAL;
	lastUR2KnownPosition	: LREAL;
	lastERRKnownPosition	: LREAL;
	lastUSERKnownPosition	: LREAL;
END_STRUCT
END_TYPE

// ---- DUTs/TYPE_MACRO.TcDUT
TYPE TYPE_MACRO :
STRUCT
	active 	: BOOL;
	mNo 	: UDINT;
	delay 	: UDINT;
END_STRUCT
END_TYPE

// ---- DUTs/TYPE_PARAMETERS.TcDUT
TYPE TYPE_PARAMETERS :
STRUCT
	(*	Nome del programma.	*)
	prgName 			: STRING[23];
	
	(*	Numero di istruzioni del programma.	*)
	sequenceCount 		: UDINT;
	
	(*	Numero assegnato alla macchina per l'identificazione, serve per collegamento in rete (opzionale).	*)
	machineNo 			: UDINT;
	
	(*	Quando arriva a zero la macchina si ferma.	*)
	pcsCounter 			: UDINT;
	
	(*	Numero di pezzi da piegare per ogni ciclo macchina.
		Il contapezzi viene decrementato di questo valore ad ogni ciclo.	*)
	pcsCycle 			: UDINT;
	
	(*	Yes: il pezzo è scaricato automaticamente a fine ciclo e le unità vanno in posizione di start del ciclo successivo.
		No 2 start: il ciclo termina con la ultime due piegature, il pezzo si deve togliere manualmente. Con uno start si portano le unità di piegatura alla posizione iniziale del ciclo successivo e con un altro start si fa ripartire il ciclo.
		No 1 start: il ciclo termina con le ultime due piegaturre, le unità di piegatura vanno automaticamente alla posizione iniziale del ciclo successvo. Il pezzo va rimosso manualmente. (si usa solo quando la posizione finale è uguale a quella inziale del ciclo successivo).	*)
	ejectMode 			: EJECT_ENUM;
	
	(*	Ritardo tra espulsione e reset ciclo (in decimi di secondo)	*)
	deltaT 				: UDINT;
	
	(*	Angolo di partenza del bracio piegatore. I minimi e massimi impostabili sono quelli impostati nei parametri macchina.
		Dopo l'azzeramento il braccio si posiziona alla quota programmata.Nome del programma.	*)
	startDegL 			: LREAL;
	
	(*	Angolo di partenza del bracio piegatore. I minimi e massimi impostabili sono quelli impostati nei parametri macchina.
		Dopo l'azzeramento il braccio si posiziona alla quota programmata.Nome del programma.	*)
	startDegR 			: LREAL;
	
	(*	Angolo di partenza per le piegature a spigolo.	*)
	startCDegL 			: LREAL;
	
	(*	Angolo di partenza per le piegature a spigolo.	*)
	startCDegR 			: LREAL;
	
	(*	Unità di movimentazione USE bilanciata o indipendente.
		Se bilanciata le unità USE si aspettatano dopo ogni istruzione.	*)
	useBalance 			: BOOL; 
	
	(*	Tabelle dei raggi varibili. *)
	radTable 			: UDINT;
	
	(*	Tabelle di elastricità. *)
	elscTable 			: UDINT;
	
	(*	 Percentuale di compensazione elasticità.	*)
	elscAdjL 			: LREAL;
	
	(*	 Percentuale di compensazione elasticità.	*)
	elscAdjR			: LREAL;
	
	(*	Tempo ciclo teorico	*)
	cycTime 			: LREAL;
	
	(*	Tempo di attrezzaggio teorico	*)
	setupTime 			: LREAL;
	
	(*	Peso del pezzo in lavorazione	*)
	pcWeight 			: LREAL;
	
	(*	Quando si raggiunde il numero di cicli macchina inserto la macchina si ferma con il bloccaggio chiuso o aperto. A seconda di Open Clamp	*)
	pcsGrpCounter 		: UDINT;
	
	(*	*)
	openClamp 			: BOOL;
	
	(*	Gradi di ritorno del braccio prima di efttuare l'inversione. Se viene messo a zero il braccio ritorna all'angolo di start.	*)
	returnDeg 			: LREAL;
	
	(*	Bloccaggio delle slitte. Se presente durante le operazioni le slitte vengono bloccate per evitare sollecitazioni alle USE.
		Funziona solo se presente nei parametri macchina.	*)
	useLockL 			: BOOL;
	
	(*	Bloccaggio delle slitte. Se presente durante le operazioni le slitte vengono bloccate per evitare sollecitazioni alle USE.
		Funziona solo se presente nei parametri macchina.	*)
	useLockR 			: BOOL;
	
	(*	Spallamento *)
	HookL 			: BOOL;
	
	(*	Spallamento *)
	HookR 			: BOOL;
	
	(*	Centering. Centratore	
		NO: Esclusione Centratore.
		TL: Centratore predisposto per la ripresa della tolleranza nei terminali del pezzo.	
		TB: Centratore predisposto per la ripresa della tolleranza in un curva (tutta la tolleranza in una curva) oppure in due curve (metà tolleranza in una curva, metà tolleranza in un'altra curva) oppure in tre o quattro curve.   *)
	centering			: CENTERING_ENUM;
	
	(*	Posizione di partenza centratore sinistro.	*)
	startL 				: LREAL;
	
	(*	Posizione di partenza centratore destro.	*)
	startR 				: LREAL;
	
	(*	Corsa rapida di avvicinamento centratore per ogni USE	*)
	inStrokeL			: LREAL;
	
	(*	Corsa rapida di avvicinamento centratore per ogni USE	*)
	inStrokeR			: LREAL;
	
	(*	Corsa massima del centratore in successione alla corsa IN STROKE   *)
	maxStrokeL			: LREAL;
	
	(*	Corsa massima del centratore in successione alla corsa IN STROKE   *)
	maxStrokeR			: LREAL;
	
		(*	Extracorsa prima della chiusura dei palpatoi.   *)
	extraL				: LREAL;
	
	(*	Extracorsa prima della chiusura dei palpatoi.   *)
	extraR				: LREAL;
	
	(*	Movimento Trasversale L.   *)
	transMovementL				: BOOL;
	
	(*	Movimento Trasversale R.   *)
	transMovementR				: BOOL;
	
	(*	Morsa del programma. TRUE: morsa normale (unita' di bloccaggio senza rotazione, motore UR2 staccato):
		il programma usa l'asse simulato UR_SIM e l'UR2 non si controlla. FALSE (default, anche con HMI che
		non lo scrivono): morsa secondo UR2Present nei parametri macchina. Cade nel padding finale: la struttura resta di 232 byte.   *)
	normalClamp					: BOOL;
	
END_STRUCT
END_TYPE

// ---- DUTs/TYPE_POSITION.TcDUT
TYPE TYPE_POSITION :
STRUCT
	active : BOOL;
	value : LREAL;
	axis : AXIS_ENUM;
END_STRUCT
END_TYPE

// ---- DUTs/TYPE_SEQUENCE.TcDUT
TYPE TYPE_SEQUENCE :
STRUCT
	active : BOOL;
	lineNo : UDINT;
	task : ARRAY[0..Size.MAX_TASK-1] OF TYPE_TASK;
END_STRUCT
END_TYPE

// ---- DUTs/TYPE_TASK.TcDUT
TYPE TYPE_TASK :
STRUCT
	active : BOOL;
	axisGroup : ARRAY[0..Size.MAX_AXIS-1] OF AXIS_ENUM;
	actions : ARRAY[0..Size.MAX_ACTION-1] OF TYPE_ACTION;
END_STRUCT
END_TYPE

// ---- Core/Cycle/E_CycleState.TcDUT
// Passi della macchina a stati del ciclo automatico (MAIN.state, Hmi.Sts.nState, Diag.Data.nState).
// I numeri sono quelli storici: compaiono nei documenti, negli allarmi ("passo 150") e nelle tracce.
// Un numero non si riusa per un passo diverso. Niente 'strict': state resta UINT e si confronta con < e >=.
// Fasce: 0-99 avvio e centraggio, 100-499 preparazione ed esecuzione, 500 fine, 600-699 abort,
//        700-799 stop e ripresa, 800-899 reset, 900-999 passaggio a manuale, 2000+ modi.
{attribute 'qualified_only'}
TYPE E_CycleState :
(
	Idle						:= 0,		// fermo, attende start
	StartChecks					:= 10,		// controlli prima di partire (lotto, azionamenti, motori, programma)

	CenteringSelect				:= 50,		// scelta del centraggio (NO/TL/TB) o posizionamento iniziale se non fatto
	Centering					:= 55,		// centraggio TL/TB in corso (FB_Centering della macchina, passo interno in Diag.Data.nSubStep)
	// 60-90: fasi del vecchio centraggio, ora dentro FB_Centering (stessi numeri). Numeri riservati.

	SeqInit						:= 110,		// azzeramento indici e sincronismi prima della prima sequenza
	SeqPrepare					:= 120,		// sequenza: gruppi e tabelle NC preparati e inviati (FB_SequenceRunner, Diag.Data.nSubStep)
	HomingPrepare				:= 122,		// homing: come SeqPrepare, con la sequenza di posizionamento iniziale
	// 130, 132, 140, 150, 200, 202, 210, 212, 400, 402: passi della vecchia preparazione, ora dentro
	// FB_SequenceRunner (E_SeqStep). Numeri riservati: non si riusano.
	SeqRun						:= 410,		// sequenza in esecuzione (RUN)
	HomingRun					:= 412,		// homing in esecuzione (INIT), poi attesa start
	WaitStartNextPiece			:= 420,		// EJECT NO 2 START: pezzo finito, attesa start

	CycleEnd					:= 500,		// fine ciclo, torna a Idle

	Abort						:= 600,		// arresto NC dei canali
	AbortDone					:= 610,		// abort concluso, avviso "reset necessario"
	WaitReset					:= 620,		// attende Reset

	Stop						:= 700,		// arresto NC per stop
	Stopped						:= 719,		// fermo, attende start (ripresa) o reset
	Resume						:= 730,		// ripresa: step-on dal RUN o reset canali
	ResumeResetTables			:= 740,		// ripresa fuori dal RUN: reset tabelle
	ResumeResetWait				:= 745,		// ripresa fuori dal RUN: attesa fine reset

	Reset						:= 800,		// reset allarmi e assi
	ResetChannels				:= 820,		// reset canali NC (non raggiunto da nessuna transizione)
	NewProgram					:= 850,		// nuovo programma dall'HMI: azzera il ciclo, poi Reset

	ToManual					:= 900,		// passaggio a manuale
	ToManualEStop				:= 905,		// passaggio a manuale: arresto NC
	ToManualClearGroups			:= 910,		// passaggio a manuale: reset gruppi
	ToManualCheckAxes			:= 915,		// passaggio a manuale: assi in errore?
	ToManualResetAxes			:= 920,		// passaggio a manuale: reset assi
	Manual						:= 2000,	// modo manuale attivo
	ToAuto						:= 2100		// passaggio ad automatico
) UINT;
END_TYPE

// ---- Core/Diag/E_CycleEndReason.TcDUT
// Perche' il ciclo automatico si e' fermato l'ultima volta (Diag.Data.eCycleEndReason).
// Si azzera allo start (passo 10).
{attribute 'qualified_only'}
{attribute 'strict'}
TYPE E_CycleEndReason :
(
	None				:= 0,	// ciclo in corso o mai partito
	PieceDone			:= 1,	// pezzo finito, il ciclo continuo riparte (o aspetta lo start con EJECT NO 2 START)
	SingleCycle			:= 2,	// pezzo finito in ciclo singolo
	BatchCompleted		:= 3,	// lotto completato (pcsCounter)
	NewProgram			:= 4,	// e' arrivato un nuovo programma: ciclo chiuso a fine pezzo
	UnknownEjectMode	:= 5,	// modo di espulsione sconosciuto (es. il vecchio EJECT 3)
	StartRefused		:= 6,	// start rifiutato nei controlli del passo 10 (vedi allarmi 63-66 e 90)
	Stopped				:= 7,	// stop dell'operatore
	Aborted				:= 8,	// abort per allarme
	ManualMode			:= 9	// passaggio a manuale
) UINT;
END_TYPE

// ---- Core/Diag/ST_DiagEvent.TcDUT
// Un cambio di passo del ciclo, con la fotografia dei canali in quel momento.
TYPE ST_DiagEvent :
STRUCT
	nIndex			: UDINT;	// progressivo dall'avvio del PLC (1 = primo evento)
	nTime			: ULINT;	// F_GetSystemTime: FILETIME, 100 ns dal 1/1/1601 UTC
	nFromState		: UINT;		// passo lasciato (E_CycleState)
	nToState		: UINT;		// passo raggiunto (E_CycleState)
	nSeqIdx			: UINT;		// sequenza corrente
	aLineNo			: ARRAY[0..Core_Param.MAX_CHANNEL-1] OF UDINT;	// riga del programma per canale (M135)
	aMFunc			: ARRAY[0..Core_Param.MAX_CHANNEL-1] OF UINT;	// funzione M richiesta e non ancora concessa, 0 = nessuna
	nAlarmId		: UINT;		// allarme memorizzato dall'evento precedente, 0 = nessuno
	nAlarmInfo		: UDINT;	// dettaglio di quell'allarme
END_STRUCT
END_TYPE

// ---- Core/Diag/ST_ChannelDiag.TcDUT
// Stato di un canale NC visto dal ciclo.
TYPE ST_ChannelDiag :
STRUCT
	bUsed			: BOOL;		// la sequenza in esecuzione ha un task su questo canale
	bDone			: BOOL;		// il canale ha finito la sua parte della sequenza
	bMWaiting		: BOOL;		// il canale chiede una funzione M e il PLC non l'ha ancora concessa
	nMFunc			: UINT;		// funzione M richiesta (0 = nessuna richiesta)
	tMWait			: TIME;		// da quanto aspetta la concessione
	nLineNo			: UDINT;	// riga del programma (M135)
	nItpState		: UDINT;	// stato dell'interprete NC (ItpGetStateInterpreter)
END_STRUCT
END_TYPE

// ---- Core/Diag/ST_Diag.TcDUT
// Diagnosi del ciclo letta dall'HMI in un solo blocco (GVL Diag.Data).
TYPE ST_Diag :
STRUCT
	nState			: UINT;					// passo attuale (E_CycleState)
	nPrevState		: UINT;					// passo precedente
	tInState		: TIME;					// da quanto il ciclo e' nel passo attuale
	nSeqIdx			: UINT;					// sequenza corrente (0 = prima)
	nSeqCount		: UINT;					// sequenze attive nel programma caricato
	nSubStep		: UINT;					// passo interno del FB al lavoro: centraggio (E_CenteringStep) o sequenza (E_SeqStep)
	eCycleEndReason	: E_CycleEndReason;		// perche' il ciclo si e' fermato l'ultima volta
	aChannel		: ARRAY[0..Core_Param.MAX_CHANNEL-1] OF ST_ChannelDiag;
	nEventCount		: UDINT;				// eventi registrati dall'avvio; l'ultimo e' aEvent[(nEventCount-1) MOD DIAG_EVENTS]
	aEvent			: ARRAY[0..Core_Param.DIAG_EVENTS-1] OF ST_DiagEvent;
	stLastAbort		: ST_DiagEvent;			// l'ultimo ingresso in abort, conservato anche quando lo storico gira
END_STRUCT
END_TYPE

// ---- Core/Valves/ST_Valve.TcDUT
// Una valvola (attuatore pneumatico) della macchina: le sue uscite e le sue conferme.
// I puntatori li assegna la configurazione della macchina a ogni ciclo (FB_MachineConfig), cosi' restano
// validi anche dopo un online change. Un feedback senza sensore puo' puntare all'uscita stessa.
TYPE ST_Valve :
STRUCT
	sName			: STRING(23);			// nome per HMI e diagnosi
	eType			: OUTPUT_ENUM;			// MONOSTABLE: solo pSet; BISTABLE: pSet e pReset
	pSet			: POINTER TO BOOL;		// uscita lato "set" (per la monostabile l'unica uscita)
	pReset			: POINTER TO BOOL;		// uscita lato "reset" (0 per la monostabile)
	pFbSet			: POINTER TO BOOL;		// conferma di fine corsa lato set
	pFbReset		: POINTER TO BOOL;		// conferma di fine corsa lato reset
END_STRUCT
END_TYPE

// ---- Core/Sync/E_MFuncKind.TcDUT
// Cosa fa il PLC quando un canale NC chiede una funzione M (handshake).
{attribute 'qualified_only'}
{attribute 'strict'}
TYPE E_MFuncKind :
(
	Nop			:= 0,	// concessa subito
	Valve		:= 1,	// muove una valvola e aspetta la conferma (timeout, post-delay): SetMacro
	ValveDirect	:= 2,	// scrive le uscite della valvola e concede subito, senza conferma
	Sync		:= 3,	// sincronismo tra canali: flag a maschera (set/clear in attesa, condizione, set/clear alla concessione)
	WaitH		:= 4,	// attesa di H millisecondi (parametro H della riga)
	LineNo		:= 5,	// numero di riga del programma nel parametro H
	WaitStart	:= 6	// attende lo start dell'operatore (passo-passo)
) UINT;
END_TYPE

// ---- Core/Sync/E_MFuncOnError.TcDUT
// Cosa succede se la valvola di una funzione M non conferma entro il timeout.
{attribute 'qualified_only'}
{attribute 'strict'}
TYPE E_MFuncOnError :
(
	Abort		:= 0,	// allarme della funzione (Info = numero M) e abort del ciclo
	Grant		:= 1,	// la funzione viene concessa lo stesso, senza allarme
	Ignore		:= 2	// nessuna reazione: il canale resta in attesa (solo per valvole la cui conferma e' l'uscita stessa)
) UINT;
END_TYPE

// ---- Core/Sync/ST_MFuncDef.TcDUT
// Una funzione M su un canale: una riga della tabella che FB_MFuncDispatcher esegue.
// Si costruisce con F_MValve, F_MValveDirect, F_MSync, F_MSimple.
TYPE ST_MFuncDef :
STRUCT
	nChannel			: UINT;				// canale NC (0 .. Core_Param.MAX_CHANNEL-1)
	nMFunc				: UINT;				// numero della funzione M
	eKind				: E_MFuncKind;

	// Valve / ValveDirect
	nValve				: UINT;				// indice nella tabella delle valvole
	eAction				: OUTPUT_ACTION_ENUM;	// SET o RESET
	tTimeout			: TIME;				// conferma attesa al massimo per...
	tPostDelay			: TIME;				// attesa dopo la conferma
	bPostDelayFromH		: BOOL;				// il post-delay e' il parametro H della riga (ms)
	nAlarmId			: UINT;				// allarme se la conferma non arriva (Info = numero M)
	eOnError			: E_MFuncOnError;
	nInterlock			: UINT;				// 0 = nessuno; altrimenti la valvola parte solo con aInterlock[nInterlock] = TRUE

	// Sync (bit di un DWORD di flag comune ai canali)
	dwSetWhileWaiting	: DWORD;			// bit messi a 1 a ogni ciclo mentre la funzione e' richiesta
	dwClearWhileWaiting	: DWORD;			// bit messi a 0 a ogni ciclo mentre la funzione e' richiesta
	dwWaitSet			: DWORD;			// condizione: questi bit tutti a 1...
	dwWaitClear			: DWORD;			// ...e questi tutti a 0
	dwSetOnGrant		: DWORD;			// bit messi a 1 alla concessione
	dwClearOnGrant		: DWORD;			// bit messi a 0 alla concessione

	nWaitAlarmId		: UINT;				// allarme di time-out mentre la condizione (sync o interlock) non e' soddisfatta; 0 = nessun time-out
END_STRUCT
END_TYPE

// ---- Machine/E_Valve.TcDUT
// Valvole di Aut260045: indice in Mach.aValve. Una valvola nuova: un valore qui, poi le sue uscite e
// conferme in FB_MachineConfig e le sue funzioni M nella tabella. Niente 'strict': e' un indice.
{attribute 'qualified_only'}
TYPE E_Valve :
(
	ErLeft			:= 1,	// testa ER SX fuori/dentro (M40/M41)
	UseLeftUp		:= 2,	// movimento trasversale ER SX su/giu' (M44/M45, diretto M54/M55)
	SupportLeft		:= 3,	// spallamento SX (M50/M51)
	EpLeftBend		:= 4,	// EP SX trazione (M70/M74), monostabile
	EpLeftOut		:= 5,	// EP SX estrazione (M72/M73)
	ErRight			:= 6,	// testa ER DX fuori/dentro (M42/M43)
	UseRightUp		:= 7,	// movimento trasversale ER DX su/giu' (M46/M47, diretto M56/M57)
	SupportRight	:= 8,	// spallamento DX (M48/M49)
	EpRightBend		:= 9,	// EP DX trazione (M70/M74), monostabile
	EpRightOut		:= 10,	// EP DX estrazione (M72/M73)
	Clamp			:= 11,	// morsa chiusa/aperta (M100/M101)
	Eject			:= 12,	// espulsore (M102/M103)
	CenteringLeftUp		:= 13,	// centratore SX su/giu' (pulsante del volantino)
	CenteringRightUp	:= 14,	// centratore DX su/giu' (pulsante del volantino)
	// Solo comandi manuali (test uscite dell'HMI); il ciclo le muove direttamente da I/O.
	CenteringUp			:= 15,	// centratori su/giu'
	CenteringClamp		:= 16,	// bloccaggio centratori, monostabile
	CenteringOut		:= 17,	// estrazione supporto centraggio, monostabile
	CenteringPiece1		:= 18,	// palpatore pezzo 1, monostabile
	CenteringPiece2		:= 19,
	CenteringPiece3		:= 20,
	CenteringPiece4		:= 21,
	CenteringAir1		:= 22,	// esclusione aria centratore 1, monostabile
	CenteringAir2		:= 23,
	CenteringAir3		:= 24,
	CenteringAir4		:= 25
) UINT;
END_TYPE

// ---- Core/Nc/ST_AxisCfg.TcDUT
// Come un asse dei programmi (valore di AXIS_ENUM in ProgramDB) entra nelle tabelle NC.
// Indice in Mach.aAxisCfg = valore di AXIS_ENUM. Un asse nuovo (es. trascinamento): una riga in FB_MachineConfig.
TYPE ST_AxisCfg :
STRUCT
	bDefined				: BOOL;			// riga configurata
	sName					: STRING(23);	// nome per HMI e diagnosi
	fSpeedScale				: LREAL;		// fVelo della riga NC = velocita' del programma * fSpeedScale
	bCenteringCorrection	: BOOL;			// alla quota si somma la correzione del centraggio TB (assi USE)
	bTargetZero				: BOOL;			// asse simulato: la quota in tabella e' sempre 0
	// Movimento manuale e servizio (FB_AxisModule)
	nMpgSelector			: UINT;			// posizione del selettore del volantino che muove l'asse (0 = nessuna)
	fJogVelocity			: LREAL;
	fJogAcceleration		: LREAL;
	fJogDeceleration		: LREAL;		// 0 = default di MC_Jog
	fJogJerk				: LREAL;
	bSoEReset				: BOOL;			// azionamento SoE reale (FB_SoEReset)
	nCalibrationAlarmId		: UINT;			// allarme per calibrazione fallita (E_Alarm della macchina)
	nLimitsAlarmId			: UINT;			// allarme per scrittura limiti fallita
	// Aggiornati dalla macchina a ogni ciclo (FB_MachineConfig)
	nNcAxisId				: UDINT;		// ID dell'asse NC (per i gruppi di interpolazione)
	fActPos					: LREAL;		// posizione attuale (punto di partenza delle tabelle)
	fActVelo				: LREAL;
	nErrorCode				: UDINT;
	bDisabled				: BOOL;
	bMoving					: BOOL;
END_STRUCT
END_TYPE

// ---- Core/Nc/E_SeqCmd.TcDUT
// Cosa il ciclo chiede a FB_SequenceRunner in questo ciclo PLC. Un comando diverso dal precedente riparte da capo.
{attribute 'qualified_only'}
{attribute 'strict'}
TYPE E_SeqCmd :
(
	None		:= 0,	// niente: solo le chiamate di servizio dei FB dei gruppi
	Prepare		:= 1,	// prepara la sequenza pSequence e la invia ai canali
	Run			:= 2,	// sequenza in esecuzione: legge la fine dei canali
	ResetTables	:= 3	// reset delle tabelle e dei canali dopo uno stop fuori dal RUN
) UINT;
END_TYPE

// ---- Core/Nc/E_SeqStep.TcDUT
// Passo interno di FB_SequenceRunner (Diag.Data.nSubStep). Tra parentesi i vecchi passi del ciclo
// (sequenza / homing) che il passo sostituisce.
{attribute 'qualified_only'}
TYPE E_SeqStep :
(
	Idle			:= 0,
	ClearGroups		:= 10,	// reset gruppi di interpolazione (120 / 122)
	BuildGroups		:= 20,	// costruzione gruppi (130 / 132)
	TableReset		:= 30,	// reset tabelle (150 / 140)
	TableStart		:= 40,	// GeoStart dalle posizioni attuali (200 / 202)
	TableFill		:= 50,	// righe di movimento e funzioni M (210 / 212)
	TableFeed		:= 60,	// invio delle tabelle ai canali (400 / 402)
	Ready			:= 100,	// tabelle inviate: la sequenza puo' girare
	Running			:= 200,	// sequenza in esecuzione (410 / 412)
	Resetting		:= 300,	// reset tabelle e canali (740 / 745)
	ResetDone		:= 310,
	Error			:= 900	// errore: vedi eErrorStep e nErrorId
) UINT;
END_TYPE

// ---- Machine/E_CenteringStep.TcDUT
// Passi di FB_Centering (Diag.Data.nSubStep durante il centraggio). Stessi numeri dei vecchi passi del ciclo.
{attribute 'qualified_only'}
TYPE E_CenteringStep :
(
	Idle				:= 0,
	ClearGroups			:= 55,	// reset dei gruppi NC per i movimenti PTP delle USE
	ApproachPrepare		:= 60,	// calcolo della corsa rapida IN STROKE
	Approach			:= 61,	// corsa rapida di avvicinamento
	ApproachCheck		:= 62,	// pezzo gia' presente prima della ricerca?
	SearchPrepare		:= 64,	// calcolo della corsa MAX STROKE
	Search				:= 65,	// ricerca dei pezzi sui sensori del centratore
	PieceClamp			:= 67,	// pezzo trovato: arresto e chiusura del palpatore
	StopAxes			:= 72,	// tutti i pezzi trovati: arresto USE
	StopDelay			:= 73,	// attesa chiusura palpatori
	Clamp				:= 74,	// chiusura morsa e calcolo della corsa EXTRA
	Extra				:= 76,	// corsa EXTRA
	ResetUnits			:= 78,	// risalita dei centratori
	Done				:= 80,	// finito
	Failed				:= 90,	// pezzo gia' presente o non trovato
	Error				:= 600	// errore NC
) UINT;
END_TYPE

// ---- Core/Nc/E_NcChannelCmd.TcDUT
// Comando a tutti i canali NC insieme (FB_NcChannels).
{attribute 'qualified_only'}
{attribute 'strict'}
TYPE E_NcChannelCmd :
(
	None		:= 0,
	EStop		:= 1,	// arresto controllato dei canali (ItpEStopEx): stop e abort
	StepOn		:= 2,	// ripartenza dal punto di arresto (ItpStepOnAfterEStopEx): ripresa dal RUN
	Reset		:= 3	// reset dei canali (ItpResetEx2)
) UINT;
END_TYPE

// ---- Core/Axes/E_AxisAlarm.TcDUT
// Allarme chiesto da FB_AxisModule in questo ciclo; il numero lo sceglie la macchina (ST_AxisCfg).
{attribute 'qualified_only'}
{attribute 'strict'}
TYPE E_AxisAlarm :
(
	None			:= 0,
	Calibration		:= 1,	// homing, lettura/scrittura offset o datum di sicurezza falliti (Info = ErrorID, 0 per il datum)
	Limits			:= 2	// scrittura dei limiti software fallita (Info = ErrorID)
) UINT;
END_TYPE

// ---- Core/Hmi/E_HmiCommand.TcDUT
// Comandi discreti dell'HMI (Hmi.Cmd.eCommand). Ogni comando ha un numero di sequenza: il PLC lo esegue una
// volta e risponde in Hmi.Sts.nCmdAck / eCmdResult. Un numero non si riusa per un comando diverso.
{attribute 'qualified_only'}
TYPE E_HmiCommand :
(
	None				:= 0,
	Start				:= 1,	// start ciclo (come il pulsante)
	Stop				:= 2,	// stop ciclo
	Reset				:= 3,	// reset allarmi e ciclo
	MotorsOn			:= 4,
	MotorsOff			:= 5,
	ProgramLoaded		:= 6,	// ProgramDB scritto: nuovo programma (azzera ciclo e contapezzi)
	WriteParameters		:= 7,	// Hmi.Param scritto: copia nei parametri macchina e scrittura dei limiti assi
	Calibrate			:= 8,	// calibrazione dell'asse nAxis; bFlag = usa la quota fValue, altrimenti la quota standard
	SetCount			:= 9	// contapezzi = nValue
) UINT;
END_TYPE

// ---- Core/Hmi/E_HmiResult.TcDUT
// Risposta del PLC a un comando (Hmi.Sts.eCmdResult).
{attribute 'qualified_only'}
TYPE E_HmiResult :
(
	None				:= 0,	// nessun comando ancora
	Accepted			:= 1,	// eseguito (l'esito del ciclo si legge negli stati e negli allarmi)
	Rejected			:= 2,	// non ammesso adesso (es. calibrazione con il ciclo in corso)
	UnknownCommand		:= 3,
	InvalidArgument		:= 4	// asse o valore fuori dai limiti
) UINT;
END_TYPE

// ---- Core/Hmi/ST_HmiCmd.TcDUT
// Comando dell'HMI (HMI -> PLC). L'HMI scrive i campi e per ultimo incrementa nSeq.
TYPE ST_HmiCmd :
STRUCT
	nSeq			: UDINT;		// cambia a ogni nuovo comando
	eCommand		: E_HmiCommand;
	nAxis			: UINT;			// asse (indice di Hmi.Cfg.aAxis) per Calibrate
	nValue			: DINT;			// valore intero (SetCount)
	fValue			: LREAL;		// valore reale (quota di Calibrate)
	bFlag			: BOOL;			// opzione (Calibrate: usa fValue)
END_STRUCT
END_TYPE

// ---- Core/Hmi/ST_HmiLive.TcDUT
// Ingressi continui dell'HMI (HMI -> PLC, scritti a ogni scambio).
TYPE ST_HmiLive :
STRUCT
	nWatchdog		: UDINT;		// l'HMI lo incrementa almeno ogni secondo: se resta fermo 3 s l'interfaccia v2 e' scollegata
	fOverride		: LREAL;		// override velocita' 0-100 %
	bLoopMode		: BOOL;			// ciclo continuo (FALSE = pezzo singolo)
	nNcMode			: UINT;			// modo dell'interprete NC (E_ItpSingleBlockMode: 0 = continuo)
	nJogAxis		: UINT;			// asse in jog (indice di Hmi.Cfg.aAxis), 0 = nessuno; solo in manuale a ciclo fermo
	nJogDirection	: INT;			// 1 avanti, -1 indietro, 0 fermo
	bForceOutputs	: BOOL;			// test uscite: le valvole seguono aValveForce
	aValveForce		: ARRAY[1..Core_Param.MAX_VALVE] OF BOOL;	// uscita "set" voluta per valvola (la "reset" e' il contrario)
END_STRUCT
END_TYPE

// ---- Core/Hmi/ST_HmiAxisParam.TcDUT
// Parametri macchina di un asse scritti dall'HMI (Hmi.Param.aAxis, applicati con il comando WriteParameters).
TYPE ST_HmiAxisParam :
STRUCT
	bPresent		: BOOL;
	bCalibrated		: BOOL;
	bCheckDone		: BOOL;			// posizione verificata dopo l'accensione
	fUpperLimit		: LREAL;		// finecorsa software massimo
	fLowerLimit		: LREAL;		// finecorsa software minimo
END_STRUCT
END_TYPE

// ---- Core/Hmi/ST_HmiParam.TcDUT
// Parametri macchina scritti dall'HMI (HMI -> PLC); diventano effettivi con il comando WriteParameters.
TYPE ST_HmiParam :
STRUCT
	bEnableSirenOverride	: BOOL;
	aAxis					: ARRAY[1..Core_Param.MAX_AXIS] OF ST_HmiAxisParam;
END_STRUCT
END_TYPE

// ---- Core/Hmi/ST_HmiNamedItem.TcDUT
// Voce di un elenco di configurazione (assi, valvole, ingressi) per costruire le pagine dell'HMI.
TYPE ST_HmiNamedItem :
STRUCT
	bDefined		: BOOL;
	sName			: STRING(23);
	nOption			: UINT;			// assi: selettore del volantino; valvole: 1 = bistabile; ingressi: 0
END_STRUCT
END_TYPE

// ---- Core/Hmi/ST_HmiCfg.TcDUT
// Configurazione della macchina per l'HMI (PLC -> HMI): si legge alla connessione.
// Le pagine dei comandi manuali e i controlli di capacita' del programma si costruiscono da qui.
TYPE ST_HmiCfg :
STRUCT
	nInterfaceVersion	: UINT;		// 2
	sMachine			: STRING(23);	// identificativo della macchina
	nMaxSequence		: UINT;		// capacita' di ProgramDB (Size.MAX_*)
	nMaxTask			: UINT;
	nMaxAction			: UINT;
	nMaxPosition		: UINT;
	nMaxMacro			: UINT;
	nMaxAxisInGroup		: UINT;
	nChannels			: UINT;
	aAxis				: ARRAY[1..Core_Param.MAX_AXIS] OF ST_HmiNamedItem;	// indice = AXIS_ENUM
	aValve				: ARRAY[1..Core_Param.MAX_VALVE] OF ST_HmiNamedItem;
	aInput				: ARRAY[1..Core_Param.MAX_INPUT] OF ST_HmiNamedItem;
END_STRUCT
END_TYPE

// ---- Core/Hmi/ST_HmiAxisSts.TcDUT
// Stato di un asse per l'HMI.
TYPE ST_HmiAxisSts :
STRUCT
	fActPos			: LREAL;
	fActVelo		: LREAL;
	nErrorCode		: UDINT;
	bEnabled		: BOOL;		// alimentato
	bMoving			: BOOL;
	bInUse			: BOOL;		// usato dalla macchina (UR2 o UR_SIM secondo la morsa)
	nCalibrationStep: UINT;		// 0 = nessuna calibrazione in corso
	bCalibrated		: BOOL;		// impulso a calibrazione finita
	bLimitsBusy		: BOOL;
	fLastKnownPos	: LREAL;	// ultima posizione salvata (persistente)
END_STRUCT
END_TYPE

// ---- Core/Hmi/ST_HmiValveSts.TcDUT
// Stato di una valvola per l'HMI.
TYPE ST_HmiValveSts :
STRUCT
	bSet			: BOOL;		// uscita "set"
	bReset			: BOOL;		// uscita "reset" (bistabile)
	bFbSet			: BOOL;		// conferma lato set
	bFbReset		: BOOL;		// conferma lato reset
END_STRUCT
END_TYPE

// ---- Core/Hmi/ST_HmiSts.TcDUT
// Stato della macchina per l'HMI (PLC -> HMI): un solo blocco letto a ogni scambio.
TYPE ST_HmiSts :
STRUCT
	nCmdAck			: UDINT;		// nSeq dell'ultimo comando trattato
	eCmdResult		: E_HmiResult;
	bConnected		: BOOL;			// il PLC vede vivo il watchdog v2
	nState			: UINT;			// passo del ciclo (E_CycleState)
	nSubStep		: UINT;			// passo interno (Diag.Data.nSubStep)
	eCycleEndReason	: E_CycleEndReason;
	bIdle			: BOOL;
	bCanExecute		: BOOL;
	bRunning		: BOOL;
	bStopped		: BOOL;
	bAborted		: BOOL;
	bHomingDone		: BOOL;
	bManualMode		: BOOL;
	bAutoMode		: BOOL;
	bMotorsOn		: BOOL;			// tutti gli azionamenti in uso abilitati
	bMotorsEnable	: BOOL;			// nessun azionamento in errore
	bLimitsWriting	: BOOL;
	bWriteParametersDone : BOOL;
	nCount			: UINT;			// contapezzi
	nSeqIdx			: UINT;
	sProgramName	: STRING(23);
	aLineNo			: ARRAY[0..Core_Param.MAX_CHANNEL-1] OF UDINT;
	aChannelDone	: ARRAY[0..Core_Param.MAX_CHANNEL-1] OF BOOL;
	nMpgSelector	: DINT;
	nMpgSpeed		: DINT;
	aAxis			: ARRAY[1..Core_Param.MAX_AXIS] OF ST_HmiAxisSts;
	aValve			: ARRAY[1..Core_Param.MAX_VALVE] OF ST_HmiValveSts;
	aInput			: ARRAY[1..Core_Param.MAX_INPUT] OF BOOL;
	aAlarmActive	: ARRAY[0..Core_Param.MAX_ALARM] OF BOOL;		// copia di Alarms.Active
	aAlarmInfo		: ARRAY[0..Core_Param.MAX_ALARM] OF UDINT;	// copia di Alarms.Info
END_STRUCT
END_TYPE

// ---- Core/Valves/ST_Input.TcDUT
// Un ingresso (sensore) della macchina mostrato all'HMI. Il puntatore lo assegna FB_MachineConfig a ogni ciclo.
TYPE ST_Input :
STRUCT
	sName			: STRING(23);
	pInput			: POINTER TO BOOL;
END_STRUCT
END_TYPE

// ---- GVLs/Alarms.TcGVL
// Allarmi macchina: un BOOL per allarme, indicizzato con E_Alarm (l'indice 0 non si usa).
// - allarmi a livello: ricalcolati a ogni ciclo in MAIN.AlarmManager, rientrano da soli;
// - allarmi memorizzati: RaiseAlarm(), restano attivi fino al Reset (ClearAlarms() nello stato 800).
// L'HMI legge Active e Info via ADS a ogni scambio.
{attribute 'qualified_only'}
VAR_GLOBAL
	Active					: ARRAY[0..Size.MAX_ALARM] OF BOOL;		// allarme attivo
	Info					: ARRAY[0..Size.MAX_ALARM] OF UDINT;	// dettaglio: ErrorID NC/azionamento, numero funzione M, 0 = nessuno
	Count					: UINT;		// allarmi attivi
	CountBlocking			: UINT;		// allarmi attivi esclusi avvisi (63-66, 90-99): accendono la torretta rossa e spengono la spia start
	StartBlockedByCabinet	: BOOL;		// almeno un allarme quadro elettrico (40-45) attivo: lo start viene rifiutato
	// Per la diagnosi (Diag.Data.aEvent): ultimo allarme memorizzato con RaiseAlarm che non era gia' attivo.
	RaisedCount				: UDINT;	// cresce a ogni nuovo allarme memorizzato
	LastRaisedId			: UINT;
	LastRaisedInfo			: UDINT;
END_VAR

// ---- GVLs/Calibration.TcGVL
{attribute 'qualified_only'}
VAR_GLOBAL
	// Quote standard usate da MC_Home quando l'override ADS non e abilitato.
	ERLHomePosition		: LREAL := 0;
	USELHomePosition	: LREAL := 1400;
	URHomePosition		: LREAL := 0;
	ERRHomePosition		: LREAL := 0;
	USERHomePosition	: LREAL := 1400;
END_VAR

// ---- GVLs/IO.TcGVL
{attribute 'qualified_only'}
VAR_GLOBAL
 	erLeftIn				AT %I* : BOOL;
	erLeftOut				AT %I* : BOOL;
	useLeftUp 				AT %I* : BOOL;
	useLeftDown 			AT %I* : BOOL;
	erRightIn 				AT %I* : BOOL;
	erRightOut 				AT %I* : BOOL;
	useRighttUp				AT %I* : BOOL;
	useRightDown			AT %I* : BOOL;
	centering1LeftIn		AT %I* : BOOL;
	centering2LeftIn		AT %I* : BOOL;
	centering3LeftIn		AT %I* : BOOL;
	centering4LeftIn		AT %I* : BOOL;
	//selectorSwitchAut1Op 	AT %I* : BOOL;
	//selectorSwitchAut2Op 	AT %I* : BOOL;
	//selectorSwitchAut 		AT %I* : BOOL;
	//selectorSwitchMan		AT %I* : BOOL;
	doorRightClosed			AT %I* : BOOL;
	doorLeftClosed			AT %I* : BOOL;
	epLeftIn				AT %I* : BOOL;
	epLeftOut				AT %I* : BOOL;
	epLeftBendDown			AT %I* : BOOL;
	epLeftBendUp			AT %I* : BOOL;
	epRightIn				AT %I* : BOOL;
	epRightOut				AT %I* : BOOL;
	epRightBendDown			AT %I* : BOOL;
	epRightBendUp			AT %I* : BOOL;
	clampIn					AT %I* : BOOL;
	bimanualStop			AT %I* : BOOL;
	bimanualOpenClamp		AT %I* : BOOL;
	fixedClampEncode		AT %I* : BOOL;
	mobileClampEncode		AT %I* : BOOL;
	clampOpen				AT %I* : BOOL;
	fuseAlarm				AT %I* : BOOL;
	leftAxisMagnetTrip		AT %I* : BOOL;
	rightAxisMagnetTrip		AT %I* : BOOL;
	ur2MagnetTrip			AT %I* : BOOL;
	chillerAlarm			AT %I* : BOOL;
	chillerMagnetTrip		AT %I* : BOOL;
	pressureSwMinPressure	AT %I* : BOOL;
	cabinetThermostat		AT %I* : BOOL;
	
	fuseReset				AT %Q* : BOOL;
	chillerEnabled			AT %Q* : BOOL;
	turretRed				AT %Q* : BOOL;
	turretYellow			AT %Q* : BOOL;
	turretGreen				AT %Q* : BOOL;
	turretSiren				AT %Q* : BOOL;
	smc1 					AT %Q* : ARRAY[0..3] OF USINT;
	smc2 					AT %Q* : ARRAY[0..3] OF USINT;
	
	useLeftUpSet 			: BOOL;
	useLeftUpReset 			: BOOL;
	useRightUpSet 			: BOOL;
	useRightUpReset 		: BOOL;
	
	erLeftOutSet 			: BOOL;
	erLeftOutReset 			: BOOL;
	erRightOutSet 			: BOOL;
	erRightOutReset 		: BOOL;
	
	supportLeftOutSet 		: BOOL;
	supportLeftOutReset 	: BOOL;
	supportRightOutSet 		: BOOL;
	supportRightOutReset	: BOOL;
	
	clampClosedSet 			: BOOL;
	clampClosedReset		: BOOL;
	
	clampEjectSet 			: BOOL;
	clampEjectReset			: BOOL;
	
	centringClamp1Left 		: BOOL;
	centringClamp2Left 		: BOOL;
	centringClamp3Left 		: BOOL;
	centringClamp4Left 		: BOOL;
	
	centeringLeft1Set 		: BOOL;
	centeringLeft2Set 		: BOOL;
	centeringLeft3Set 		: BOOL;
	centeringLeft4Set 		: BOOL;
	
	centeringLeft1Reset 	: BOOL;
	centeringLeft2Reset 	: BOOL;
	centeringLeft3Reset 	: BOOL;
	centeringLeft4Reset 	: BOOL;
		
	centeringRight1Set 		: BOOL;
	centeringRight2Set 		: BOOL;
	centeringRight3Set 		: BOOL;
	centeringRight4Set 		: BOOL;
	
	centeringRight1Reset 	: BOOL;
	centeringRight2Reset 	: BOOL;
	centeringRight3Reset 	: BOOL;
	centeringRight4Reset 	: BOOL;
	
	centringClampSet		: BOOL;
	
	centringLeftUpSet 		: BOOL;
	centringLeftUpReset 	: BOOL;
	
	centringRightUpSet 		: BOOL;
	centringRightUpReset 	: BOOL;
	
	centeringLeftReset		: BOOL;
	centeringRightReset		: BOOL;
	
	centringSet 			: BOOL;
	centringReset 			: BOOL;
	
	centeringOutSet			: BOOL; //Estrazione verso destra supporto bloccaggio / centraggio
	
	Pc1CenteringLock		: BOOL;
	Pc2CenteringLock		: BOOL;
	
	epLeftOutSet			: BOOL;
	epLeftOutReset			: BOOL;
	epLeftBend				: BOOL;
	
	epRightOutSet			: BOOL;
	epRightOutReset			: BOOL;
	epRightBend				: BOOL;
	
	spiaPulsanteStart 		AT %Q* : BOOL;
	spiaPulsanteStop 		AT %Q* : BOOL;
END_VAR

// ---- GVLs/Machine.TcGVL
{attribute 'qualified_only'}
VAR_GLOBAL PERSISTENT
	parametersRx : TYPE_MACHINE_RX;
	parametersTx : TYPE_MACHINE_TX;
END_VAR

// ---- GVLs/ProgramDB.TcGVL
{attribute 'qualified_only'}
VAR_GLOBAL
	parameters	: TYPE_PARAMETERS;
	homing		: TYPE_SEQUENCE;
	sequence	: ARRAY[0..Size.MAX_SEQUENCE-1] OF TYPE_SEQUENCE;
	prgState	: PRGSTATE_ENUM;
END_VAR

// ---- GVLs/Safety.TcGVL
{attribute 'qualified_only'}
VAR_GLOBAL
	Run 				AT %Q* : BOOL;
	Ack 				AT %Q* : BOOL;
	ModuleFault         AT %Q* : BOOL;
	
	USER_ERR_Run 		AT %Q* : BOOL;
	USER_ERR_Ack 		AT %Q* : BOOL;
	
	USEL_ERL_Run 		AT %Q* : BOOL;
	USEL_ERL_Ack 		AT %Q* : BOOL;
	
	UR_Run 				AT %Q* : BOOL;
	UR_Ack 				AT %Q* : BOOL;
	
	FBErr 				AT %I* : BOOL;
	FBRun				AT %I* : BOOL;
	ComErr 				AT %I* : BOOL;
	OutErr 				AT %I* : BOOL;
	OtherErr 			AT %I* : BOOL;
	ComStartup 			AT %I* : BOOL;
	FBDeactivate 		AT %I* : BOOL;
	InRun 				AT %I* : BOOL;
	EmergenzaResettata 	AT %I* : BOOL;
	bimanualStart		AT %I* : BOOL;
	
	USEL_ERL_FBErr			AT %I* : BOOL;
	USEL_ERL_FBRun			AT %I* : BOOL;
	USEL_ERL_ComErr 		AT %I* : BOOL;
	USEL_ERL_OutErr 		AT %I* : BOOL;
	USEL_ERL_OtherErr 		AT %I* : BOOL;
	USEL_ERL_ComStartup 	AT %I* : BOOL;
	USEL_ERL_FBDeactivate	AT %I* : BOOL;
	USEL_ERL_InRun 			AT %I* : BOOL;
		
	USER_ERR_FBErr			AT %I* : BOOL;
	USER_ERR_FBRun			AT %I* : BOOL;
	USER_ERR_ComErr 		AT %I* : BOOL;
	USER_ERR_OutErr 		AT %I* : BOOL;
	USER_ERR_OtherErr 		AT %I* : BOOL;
	USER_ERR_ComStartup 	AT %I* : BOOL;
	USER_ERR_FBDeactivate	AT %I* : BOOL;
	USER_ERR_InRun 			AT %I* : BOOL;
	
	UR_FBErr			AT %I* : BOOL;
	UR_FBRun			AT %I* : BOOL;
	UR_ComErr 			AT %I* : BOOL;
	UR_OutErr 			AT %I* : BOOL;
	UR_OtherErr 		AT %I* : BOOL;
	UR_ComStartup 		AT %I* : BOOL;
	UR_FBDeactivate		AT %I* : BOOL;
	UR_InRun 			AT %I* : BOOL;
	
	ERLDatumRequest		AT %I* : BOOL;
	ERLDatumDone		AT %I* : BOOL;
	ERLSafetyReset		AT %Q* : SINT;
	ERLDatumExecute		AT %Q* : BOOL;
	ERLCommErrorAck		AT %Q* : BOOL;
	
	ERL_STO			AT %I* : BOOL;
	ERL_SSM1		AT %I* : BOOL;
	ERL_SSM2		AT %I* : BOOL;
	ERL_SOS			AT %I* : BOOL;
	ERL_SSR			AT %I* : BOOL;
	ERL_SDI_p		AT %I* : BOOL;
	ERL_SDI_n		AT %I* : BOOL;
	ERL_Error		AT %I* : BOOL;
	
	USEL_STO		AT %I* : BOOL;
	USEL_SSM1		AT %I* : BOOL;
	USEL_SSM2		AT %I* : BOOL;
	USEL_SOS		AT %I* : BOOL;
	USEL_SSR		AT %I* : BOOL;
	USEL_SDI_p		AT %I* : BOOL;
	USEL_SDI_n		AT %I* : BOOL;
	USEL_Error		AT %I* : BOOL;
	
	ERR_STO			AT %I* : BOOL;
	ERR_SSM1		AT %I* : BOOL;
	ERR_SSM2		AT %I* : BOOL;
	ERR_SOS			AT %I* : BOOL;
	ERR_SSR			AT %I* : BOOL;
	ERR_SSR2		AT %I* : BOOL;
	ERR_SDI_p		AT %I* : BOOL;
	ERR_SDI_n		AT %I* : BOOL;
	ERR_Error		AT %I* : BOOL;
	
	USER_STO		AT %I* : BOOL;
	USER_SSM1		AT %I* : BOOL;
	USER_SSM2		AT %I* : BOOL;
	USER_SOS		AT %I* : BOOL;
	USER_SSR		AT %I* : BOOL;
	USER_SSR2		AT %I* : BOOL;
	USER_SDI_p		AT %I* : BOOL;
	USER_SDI_n		AT %I* : BOOL;
	USER_Error		AT %I* : BOOL;
	
	UR_STO		AT %I* : BOOL;
	UR_SSM1		AT %I* : BOOL;
	UR_SSM2		AT %I* : BOOL;
	UR_SOS		AT %I* : BOOL;
	UR_SSR		AT %I* : BOOL;
	UR_SDI_p		AT %I* : BOOL;
	UR_SDI_n		AT %I* : BOOL;
	UR_Error		AT %I* : BOOL;

	USELDatumRquest		AT %I* : BOOL;
	USELDatumDone		AT %I* : BOOL;
	USELSafetyReset		AT %Q* : SINT;
	USELDatumExecute	AT %Q* : BOOL;
	USELCommErrorAck	AT %Q* : BOOL;
	
	URDatumRequest		AT %I* : BOOL;
	URDatumDone			AT %I* : BOOL;
	URSafetyReset		AT %Q* : SINT;
	URDatumExecute		AT %Q* : BOOL;
	URCommErrorAck		AT %Q* : BOOL;
	
	ERRDatumRequest		AT %I* : BOOL;
	ERRDatumDone		AT %I* : BOOL;
	ERRSafetyReset		AT %Q* : SINT;
	ERRDatumExecute		AT %Q* : BOOL;
	ERRCommErrorAck		AT %Q* : BOOL;
	
	USERDatumRequest	AT %I* : BOOL;
	USERDatumDone		AT %I* : BOOL;
	USERSafetyReset		AT %Q* : SINT;
	USERDatumExecute	AT %Q* : BOOL;
	USERCommErrorAck	AT %Q* : BOOL;
	
	ResetEmergenza		AT %Q* : BOOL;
	ResetBarriere		AT %Q* : BOOL;
	PulsanteResetBarriere AT %I* : BOOL;
	PulsanteResetEmergenza AT %I* : BOOL;
	BarriereResettate      AT %I* : BOOL;
	
	SpiaPulsanteRipristinoSicurezze 	AT %Q* : BOOL;
	SpiaPulsanteRipristinoBarriere 		AT %Q* : BOOL;
	ModoSemiAuto						AT %I* : BOOL;
	ModoManuale							AT %I* : BOOL;
	ModoAuto1Op							AT %I* : BOOL;
	ModoAuto2Op							AT %I* : BOOL;
	AbilitazionePeriferiche				AT %I* : BOOL;
	
	SSR1_Enable 						AT %I* : BOOL;
	SSR2_Enable 						AT %I* : BOOL;
END_VAR

// ---- GVLs/Size.TcGVL
{attribute 'qualified_only'}
// Capacita' di ProgramDB: ogni MAX_* e' il NUMERO di elementi, gli array vanno da 0 a MAX_*-1.
// Devono restare uguali ai limiti dell'HMI (PlcSequenceBuilder): cambiarli cambia il layout ADS di ProgramDB.
VAR_GLOBAL	CONSTANT
	MAX_SEQUENCE 	: UINT := 100;
	MAX_TASK 		: UINT := 3;
	MAX_ACTION 		: UINT := 24;
	MAX_POSITION 	: UINT := 8;
	MAX_AXIS 		: UINT := 8;
	MAX_MACRO 		: UINT := 8;
	MAX_ALARM		: UINT := 255;	// ultimo indice di Alarms.Active / Alarms.Info (E_Alarm)
END_VAR

// ---- Core/Core_Param.TcGVL
// Dimensioni del Core. Quando il Core diventera' una libreria questa lista sara' la sua parameter list:
// ogni macchina la imposta senza toccare il codice del Core.
{attribute 'qualified_only'}
VAR_GLOBAL CONSTANT
	MAX_CHANNEL		: UINT := 3;	// canali NC di interpolazione (SX, DX, UR2)
	DIAG_EVENTS		: UINT := 64;	// eventi tenuti nello storico della diagnosi
	MAX_AXIS		: UINT := 16;	// assi configurabili (indice = AXIS_ENUM)
	MAX_VALVE		: UINT := 32;	// valvole configurabili
	MAX_INPUT		: UINT := 32;	// ingressi mostrati all'HMI
	MAX_ALARM		: UINT := 255;	// ultimo indice degli allarmi (uguale a Size.MAX_ALARM)
END_VAR

// ---- GVLs/Diag.TcGVL
// Diagnosi del ciclo per l'HMI: una sola lettura ADS di Diag.Data (MAIN.DiagUpdate la aggiorna a ogni ciclo).
{attribute 'qualified_only'}
VAR_GLOBAL
	Data		: ST_Diag;
END_VAR

// ---- Machine/Mach.TcGVL
// Configurazione di Aut260045 usata dal Core: valvole, funzioni M, interblocchi.
// La riempie FB_MachineConfig (MAIN.fbMachineConfig) a ogni ciclo.
{attribute 'qualified_only'}
VAR_GLOBAL CONSTANT
	MAX_VALVE		: UINT := Core_Param.MAX_VALVE;
	MAX_MFUNC		: UINT := 96;
	MAX_INTERLOCK	: UINT := 8;
	MAX_AXIS_CFG	: UINT := Core_Param.MAX_AXIS;	// valori di AXIS_ENUM configurabili (1..16)
	NC_GROUP_BASE	: UDINT := 7;	// ID NC del gruppo di interpolazione del canale 0 (canali 7, 8, 9)
	MAX_MPG_SEL		: UINT := 8;	// posizioni del selettore del volantino

	// Indici degli assi in aAxisCfg e in MAIN.aAxisMod (= valori di AXIS_ENUM)
	AX_USEL			: UINT := 1;
	AX_USER			: UINT := 2;
	AX_ERL			: UINT := 3;
	AX_ERR			: UINT := 4;
	AX_UR2			: UINT := 5;
	AX_UR_SIM		: UINT := 6;

	// Interblocchi (indice in aInterlock)
	IL_UR2_AT_ZERO	: UINT := 1;	// UR2 entro 3 gradi da zero, o UR2 non usato: l'espulsore puo' partire (M102)

	// Flag di sincronismo tra i canali (bit di MAIN.syncFlags)
	SYNC_ACK_L		: DWORD := 16#0001;	// USE SX in posizione (M62), atteso da DX (M60) e UR2 (M116)
	SYNC_ACK_R		: DWORD := 16#0002;	// USE DX in posizione (M63), atteso da SX (M61) e UR2 (M116)
	SYNC_ACK_UR2	: DWORD := 16#0004;	// riservato (azzerato da M150 sull'UR2)
	SYNC_UR2_DONE	: DWORD := 16#0008;	// UR2 in posizione (M78), atteso dalle USE (M80)
	SYNC_UR2_ACK_L	: DWORD := 16#0010;	// USE SX ha visto l'UR2 (M112), atteso dall'UR2 (M110)
	SYNC_UR2_ACK_R	: DWORD := 16#0020;	// USE DX ha visto l'UR2 (M113), atteso dall'UR2 (M110)
	SYNC_DONE_L		: DWORD := 16#0040;	// riservato (azzerato da M150 su SX)
	SYNC_DONE_R		: DWORD := 16#0080;	// riservato (azzerato da M150 su DX)
	SYNC_UR2_REQ_L	: DWORD := 16#0100;	// riservato (azzerato da M150 sull'UR2)
	SYNC_UR2_REQ_R	: DWORD := 16#0200;	// riservato (azzerato da M150 sull'UR2)
END_VAR
VAR_GLOBAL
	aAxisCfg		: ARRAY[1..Mach.MAX_AXIS_CFG] OF ST_AxisCfg;	// indice = valore di AXIS_ENUM
	aValve			: ARRAY[1..Mach.MAX_VALVE] OF ST_Valve;
	aInput			: ARRAY[1..Core_Param.MAX_INPUT] OF ST_Input;	// ingressi mostrati all'HMI (sensori)
	aMFunc			: ARRAY[1..Mach.MAX_MFUNC] OF ST_MFuncDef;
	nMFuncCount		: UINT;		// righe valide di aMFunc
	aInterlock		: ARRAY[0..Mach.MAX_INTERLOCK] OF BOOL;	// l'indice 0 non si usa (0 = nessun interblocco)
	// Pulsanti del volantino per posizione del selettore: [selettore, 1] = pulsante 1, [selettore, 2] = pulsante 3.
	// Valore = valvola (E_Valve) da commutare, 0 = nessuna.
	aMpgButton		: ARRAY[1..Mach.MAX_MPG_SEL, 1..2] OF UINT;
END_VAR

// ---- GVLs/Hmi.TcGVL
// Interfaccia HMI v2 (contratto in docs/ADS_CONTRACT_V2.md). Ogni blocco si legge o scrive con una chiamata ADS.
// E' l'unica interfaccia con l'HMI: la v1 (GVL Ads) e' stata tolta.
{attribute 'qualified_only'}
VAR_GLOBAL
	Cfg			: ST_HmiCfg;		// PLC -> HMI, alla connessione: assi, valvole, ingressi, capacita'
	Cmd			: ST_HmiCmd;		// HMI -> PLC: comando con numero di sequenza
	Live		: ST_HmiLive;		// HMI -> PLC, ciclico: watchdog, override, jog, test uscite
	Param		: ST_HmiParam;		// HMI -> PLC: parametri macchina, applicati con il comando WriteParameters
	Sts			: ST_HmiSts;		// PLC -> HMI, ciclico: stato, assi, valvole, ingressi, allarmi
END_VAR

// ---- POUs/MAIN.TcPOU
PROGRAM MAIN
VAR
//V1.10
//*******************************************************************************************************************
// Parameters
//*******************************************************************************************************************
	USEMoveSpeed				: LREAL := 200;	//Use speed during centering
	USESearchSpeed				: LREAL := 30;	//Use speed during centering research
	tMotorsOffDelay				: TIME := T#100MS;	//Time before motors off event
	channel1SafeOverride		: REAL := 10;
	channel2SafeOverride		: REAL := 10;
	channel3SafeOverride		: REAL := 10;
	uselSafeOvPosition			: LREAL := 140;
	userSafeOvPosition			: LREAL := 140;
	tSyncTimeOut				: TIME := T#15S;	//max wait on M60/61/80/102/110/112/113/116 with the cycle not progressing (manual: about 15 s)
	tStateTimeOut				: TIME := T#10S;	//max time in a technical state (NC/MC function blocks only), then StateTimeout

	urUSELMinPosition			: LREAL := 65;
	urUSERMinPosition			: LREAL := 65;
	ur2USELMinPosition			: LREAL := 95;
	ur2USERMinPosition			: LREAL := 95;
//*******************************************************************************************************************
// Bools
//*******************************************************************************************************************
	motorsOn					: BOOL;		//Motors Torque on instructions
	motorsOffTrigger			: BOOL;		//Motors off trigger
	allDrivesEnabled 			: BOOL;		//true when all drivers are enabled
	ur2InUse					: BOOL;		//true when the UR2 unit is used: UR2Present and the program does not mount the normal clamp
	ur2InUsePrev				: BOOL;		//ur2InUse already applied to the USE soft limits
	newProgramTrigger			: BOOL;		//true for one cycle when the HMI loads a new program (command ProgramLoaded)
	newProgramPending			: BOOL;		//true while the cycle reset for the new program is pending
	drivesError					: BOOL;		//true when a drive is in error state
	homingDone					: BOOL;		//true when homing done
	USELDone					: BOOL;		//true when USEL completed its instructions
	USERDone					: BOOL;
	UR2Done						: BOOL;
	USEL_UR2_Ack				: BOOL;		//acknolage of UR2 from USE
	USER_UR2_Ack				: BOOL;
	UR2_USEL_Req				: BOOL;		//achnlage request frin UR2 TO USE
	UR2_USER_Req				: BOOL;
	manualMode					: BOOL;		//true when manual mode active
	autoMode					: BOOL;		//true when auto mode active
	manualModeTrigger			: BOOL;		//trigger to switch to manual mode
	autoModeTrigger				: BOOL;		//trigger to switch to auto mode
	firstScan					: BOOL := TRUE;
	autoLoopMode				: BOOL;
	startTriggerOut				: BOOL;
	bimanualOpenClampTriggerOut	: BOOL;
	startCondition				: BOOL;
	programIdle					: BOOL;
	programCanExecute			: BOOL;
	programAborted				: BOOL;
	programStopped				: BOOL;
	programRunning				: BOOL;
	safeOverride				: BOOL;
	writeParametersEvent		: BOOL;
	writeParametersDone			: BOOL;		//last axis limits writing ended without errors (Hmi.Sts.bWriteParametersDone)
	nextSequenceActive			: BOOL;		//state 410: the sequence after seqIdx exists and is active
	stopPending					: BOOL;		//stop pressed during centering, INIT or end-of-piece wait: applied at the end of the phase
	clampClosedAtStop			: BOOL;		//clamp command when the stop was applied (state 700), restored on resume
	syncBlockedAll				: BOOL;		//every channel is done, unused or waiting for a sync: the cycle is not progressing
	stateWatchPrev				: UINT;		//state seen by the state watchdog in the previous scan
	stateIsTechnical			: BOOL;		//current state only waits for an NC/MC function block (watched by fbStateWatchdog)
	cycleEndReason				: E_CycleEndReason;	//why the automatic cycle stopped the last time (Diag.Data.eCycleEndReason)
	diagSeqIdx					: UINT;		//loop index used by DiagUpdate to count the active sequences
	diagSeqCounted				: BOOL;		//DiagUpdate has counted the sequences at least once since PLC start
	syncTaskInUse				: BOOL;
	channelDone					: ARRAY[0..2] OF BOOL;
	syncAck						: ARRAY[0..2] OF BOOL;
	syncFlags					: DWORD;	//sync flags packed for fbMFunc (bits Mach.SYNC_*), unpacked again after the call
	syncWait					: ARRAY[0..2] OF BOOL;		//channel waiting on a sync M function (or M102 with UR2 not at zero)
	bLogEntries					: ARRAY[0..2] OF BOOL;
	bMotorsOnStatus				: ARRAY[0..4] OF BOOL;
//*******************************************************************************************************************
// Uint
//*******************************************************************************************************************
	i							: UINT;
	lastState					: UINT;
	seqIdx						: UINT;
	lineNo1						: UDINT;
	lineNo2						: UDINT;
	lineNo3						: UDINT;
	state						: UINT := 0;
	count						: UINT := 0;
	alarmIdx					: UINT;		//indice per i conteggi allarmi
	udiItpState					: ARRAY[0..2] OF UDINT;
	syncWaitAlarm				: ARRAY[0..2] OF UINT;		//time-out alarm (E_Alarm) of the sync wait in progress on each channel
//*******************************************************************************************************************
// LREAL
//*******************************************************************************************************************
	MeasureL					: LREAL;
	MeasureR					: LREAL;
	ToleranceMeasure			: LREAL;
	axisOverride				: LREAL := 100;
	channel1Override			: REAL;
	channel2Override			: REAL;
	channel3Override			: REAL;
	
//*******************************************************************************************************************
// STs
//******************************************************************************************************************
	parametersRx 				: TYPE_MACHINE_RX;
	stMpgEncoder 				: ST_MpgEncoder;
	stTwoHandControl			: ST_TwoHandControl;
//*******************************************************************************************************************
// FBs
//******************************************************************************************************************
	fbSelectorOnTrigger			: R_TRIG;
	fbSelectorOffTrigger		: R_TRIG;
	fbBimanualOpenClampTrigger	: R_TRIG;
	fbCloseClampAfterCentering	: TON;
	ssrActivationDelay			: TON;
	ssr2ActivationDelay			: TON;
	waitForMove					: TON;
	USEL 						: AXIS_REF;
	ERL 						: AXIS_REF;
	USER 						: AXIS_REF;
	ERR 						: AXIS_REF;
	UR2 						: AXIS_REF;
	UR_SIM 						: AXIS_REF;
	fbMPGReadStatus				: MPG_ReadStatus;
	fbTwoHandReadStatus			: TwoHand_ReadStatus;
	fbTimerOffMotos				: ARRAY[0..4] OF TOF;
	fbSeq						: FB_SequenceRunner;	//NC groups and tables of the running sequence (prepare, run, reset)
	seqCmd						: E_SeqCmd;		//command given to fbSeq in this scan, from the cycle state
	seqAlarmId					: UINT;			//alarm (E_Alarm) for an fbSeq error during preparation
	fbCentering					: FB_Centering;		//TL/TB centering phase (cycle step Centering)
	fbNc						: FB_NcChannels;		//e-stop, step-on and reset of all NC channels
	ncCmd						: E_NcChannelCmd;	//command given to fbNc in this scan, from the cycle state
	aAxisMod					: ARRAY[1..Mach.MAX_AXIS_CFG] OF FB_AxisModule;	//one module per axis (index = AXIS_ENUM value, Mach.AX_*)
	axisInUse					: ARRAY[1..Mach.MAX_AXIS_CFG] OF BOOL;		//axis powered, jogged and reset (UR2 or UR_SIM by ur2InUse)
	resetAxesCmd				: BOOL;		//MC_Reset of the axes in use (cycle steps 800, 920), cleared every scan in InitCyclic
	axesResetDone				: BOOL;
	axesResetError				: BOOL;
	axesResetErrorId			: UDINT;
	limitsRequest				: BOOL;		//rewrite the axis limits (clamp changed)
	limitsStart					: BOOL;		//this scan starts the limits writing (HMI command or limitsRequest)
	limitsWriting				: BOOL;		//limits writing in progress: the cycle does not start
	limitsBusy					: BOOL;
	limitsFailed				: BOOL;
	limitsAxis					: UINT;		//last axis whose limits writing was started (0 = none yet)
	limitsKickAxis				: UINT;		//axis that starts its limits writing in the next scan (0 = none)
	calibrationBusy				: BOOL;		// calibrazione richiesta o in corso: impedisce l'avvio ciclo
	mpgSelector					: UINT;		//handwheel selector position
	mpgAxisSelected				: BOOL;
	mpgValve					: UINT;
	jogSelected					: BOOL;
	fbHmiWatchdog				: FB_HmiWatchdog;	//HMI alive (Hmi.Live.nWatchdog)
	fbHmiCmd					: FB_HmiCommandHandler;	//HMI commands with sequence number (Hmi.Cmd)
	hmiConnected				: BOOL;		//HMI connected: watchdog of Hmi.Live alive
	hmiStartCmd					: BOOL;
	hmiStopCmd					: BOOL;
	hmiResetCmd					: BOOL;
	hmiMotorsOnCmd				: BOOL;
	hmiMotorsOffCmd				: BOOL;
	hmiProgramLoadedCmd			: BOOL;
	hmiWriteParamsCmd			: BOOL;
	hmiStop						: BOOL;		//stop request this scan (HMI command)
	hmiReset					: BOOL;		//reset request this scan (HMI command)
	hmiOverride					: LREAL;	//speed override from the HMI (0-100)
	ncSingleBlock				: BOOL;		//NC interpreter in single-block (step) mode
	hmiForce					: BOOL;		//output test active
	valveForce					: ARRAY[1..Mach.MAX_VALVE] OF BOOL;	//output test: wanted "set" output per valve
	calibStart					: ARRAY[1..Mach.MAX_AXIS_CFG] OF BOOL;
	calibUsePos					: ARRAY[1..Mach.MAX_AXIS_CFG] OF BOOL;
	calibPos					: ARRAY[1..Mach.MAX_AXIS_CFG] OF LREAL;
	jogHmi						: BOOL;
	fbMachineConfig				: FB_MachineConfig;		//valves and M function table of this machine (Mach GVL)
	fbMFunc						: FB_MFuncDispatcher;	//executes the M functions requested by the NC channels
	fbSyncTimeOut				: ARRAY[0..2] OF TON;
	fbStateWatchdog				: TON;
	fbDiagLog					: FB_DiagLog;
	fbMFuncWait					: ARRAY[0..2] OF TON;	//time a channel has been waiting for an M function grant (diagnostics)
	fbClearGroup				: ARRAY[0..2] OF CfgReconfigGroup;
	
	fbUps 						: FB_S_UPS_BAPI; 
//*******************************************************************************************************************
// IOs
//*******************************************************************************************************************
	in_stNciToPlc AT %I* : ARRAY[0..2] OF NCTOPLC_NCICHANNEL_REF;
	out_stPlcToNci AT %Q*: ARRAY[0..2] OF PLCTONC_NCICHANNEL_REF;
END_VAR

//*******************************************************************************************************************
// init
//*******************************************************************************************************************
IF firstScan THEN
	InitOnce();
END_IF

fbUps(
    sNetID          := '',                              // '' = AmsNetId locale
    iPLCPort        := 851,                              // porta runtime PLC (851 = primo runtime)
    tTimeout        := DEFAULT_ADS_TIMEOUT,
    eUpsMode        := eSUPS_WrPersistData_Shutdown,     // salva dati persistenti poi QuickShutdown (default consigliato)
    ePersistentMode := SPDM_2PASS,                       // modo veloce, obbligatorio per la 1-sec UPS
    tRecoverTime    := T#10s
);

// Base ciclo: clock, default FB e lettura dispositivi operatore.
Clock();
InitCyclic();
fbMPGReadStatus(stMpgEncoder := stMpgEncoder);
fbTwoHandReadStatus(stTwoHandControl := stTwoHandControl);

// Ingressi esterni e consensi macchina.
HmiInputs();
SafetyManager();
InputMapping();
MotorStatusManager();
ParameterWriteManager();
DriveStatusManager();

// Configurazione della macchina per il Core (assi, valvole, funzioni M) con ID e posizioni di questo ciclo.
fbMachineConfig();

// Esecuzione programma e macro NC.
IF manualMode THEN
	Manual();
END_IF
StateMachine();
MacroManager();

// Allarmi: dopo la macchina a stati, cosi' un Reset (stato 800) non spegne per un ciclo quelli ancora presenti.
AlarmManager();

// Diagnosi: dopo tutto cio' che puo' cambiare il passo nel ciclo (macchina a stati, funzioni M, allarmi).
DiagUpdate();

// Chiamate FB che devono girare ogni ciclo.
AxisFunctionBlocks();
OutputMapping();
HmiOutputs();

ACTION AlarmManager:
// Allarmi a livello (ricalcolati a ogni ciclo) e conteggi per torretta, spia start e interblocco.
// Gli allarmi memorizzati si attivano con RaiseAlarm() e si azzerano col Reset (stato 800).

// Sicurezza
Alarms.Active[E_Alarm.EmergencyStop]			:= NOT Safety.EmergenzaResettata;
Alarms.Active[E_Alarm.DoorLeftOpen]				:= NOT IO.doorLeftClosed;
Alarms.Active[E_Alarm.DoorRightOpen]			:= NOT IO.doorRightClosed;
Alarms.Active[E_Alarm.LightCurtainNotReset]		:= NOT Safety.BarriereResettate;
Alarms.Active[E_Alarm.SafetyMainGroupError]		:= Safety.FBErr OR Safety.ComErr OR Safety.OtherErr;
Alarms.Active[E_Alarm.SafetyGroupLeftError]		:= Safety.USEL_ERL_FBErr OR Safety.USEL_ERL_ComErr OR Safety.USEL_ERL_OtherErr;
Alarms.Active[E_Alarm.SafetyGroupRightError]	:= Safety.USER_ERR_FBErr OR Safety.USER_ERR_ComErr OR Safety.USER_ERR_OtherErr;
Alarms.Active[E_Alarm.SafetyGroupUrError]		:= Safety.UR_FBErr OR Safety.UR_ComErr OR Safety.UR_OtherErr;

// Azionamenti: Info = codice errore NC dell'asse
Alarms.Active[E_Alarm.DriveErl]		:= ERL.NcToPlc.ErrorCode <> 0 AND Machine.parametersRx.ERLPresent;
Alarms.Active[E_Alarm.DriveUsel]	:= USEL.NcToPlc.ErrorCode <> 0 AND Machine.parametersRx.USELPresent;
Alarms.Active[E_Alarm.DriveUr2]		:= UR2.NcToPlc.ErrorCode <> 0 AND ur2InUse;
Alarms.Active[E_Alarm.DriveErr]		:= ERR.NcToPlc.ErrorCode <> 0 AND Machine.parametersRx.ERRPresent;
Alarms.Active[E_Alarm.DriveUser]	:= USER.NcToPlc.ErrorCode <> 0 AND Machine.parametersRx.USERPresent;
Alarms.Info[E_Alarm.DriveErl]		:= SEL(Alarms.Active[E_Alarm.DriveErl], 0, ERL.NcToPlc.ErrorCode);
Alarms.Info[E_Alarm.DriveUsel]		:= SEL(Alarms.Active[E_Alarm.DriveUsel], 0, USEL.NcToPlc.ErrorCode);
Alarms.Info[E_Alarm.DriveUr2]		:= SEL(Alarms.Active[E_Alarm.DriveUr2], 0, UR2.NcToPlc.ErrorCode);
Alarms.Info[E_Alarm.DriveErr]		:= SEL(Alarms.Active[E_Alarm.DriveErr], 0, ERR.NcToPlc.ErrorCode);
Alarms.Info[E_Alarm.DriveUser]		:= SEL(Alarms.Active[E_Alarm.DriveUser], 0, USER.NcToPlc.ErrorCode);

// Quadro elettrico: ingressi TRUE = guasto (da verificare sullo schema alla messa in servizio)
Alarms.Active[E_Alarm.FuseTripped]		:= NOT IO.fuseAlarm;
Alarms.Active[E_Alarm.BreakerLeftAxis]	:= NOT IO.leftAxisMagnetTrip;
Alarms.Active[E_Alarm.BreakerRightAxis]	:= NOT IO.rightAxisMagnetTrip;
Alarms.Active[E_Alarm.BreakerUr2]		:= NOT IO.ur2MagnetTrip;
Alarms.Active[E_Alarm.BreakerChiller]	:= NOT IO.chillerMagnetTrip;
Alarms.Active[E_Alarm.AirPressureLow]	:= NOT IO.pressureSwMinPressure;

// Avvisi
Alarms.Active[E_Alarm.ChillerAlarm]				:= IO.chillerAlarm;
Alarms.Active[E_Alarm.CabinetOverTemperature]	:= IO.cabinetThermostat;

// Conteggi. Gli avvisi (start rifiutato 63-66, avvisi 90-99) non contano come bloccanti.
Alarms.Count := 0;
Alarms.CountBlocking := 0;
FOR alarmIdx := 1 TO Size.MAX_ALARM DO
	IF Alarms.Active[alarmIdx] THEN
		Alarms.Count := Alarms.Count + 1;
		IF NOT ((alarmIdx >= E_Alarm.StartDriveError AND alarmIdx <= E_Alarm.StartCabinetAlarm) OR (alarmIdx >= 90 AND alarmIdx <= 99)) THEN
			Alarms.CountBlocking := Alarms.CountBlocking + 1;
		END_IF
	END_IF
END_FOR

Alarms.StartBlockedByCabinet := Alarms.Active[E_Alarm.FuseTripped] OR Alarms.Active[E_Alarm.BreakerLeftAxis]
	OR Alarms.Active[E_Alarm.BreakerRightAxis] OR Alarms.Active[E_Alarm.BreakerUr2]
	OR Alarms.Active[E_Alarm.BreakerChiller] OR Alarms.Active[E_Alarm.AirPressureLow];

// Allarmi "non calibrato" per asse: disabilitati (lo erano anche con la vecchia lista messaggi).
END_ACTION

ACTION AxisFunctionBlocks:
// Esegue FB assi, NCI, macro, timer e letture parametri.


// Assi: potenza, jog, reset, calibrazione, limiti nei moduli FB_AxisModule.
AxisModules();

ItpSetOverridePercent(fOverridePercent:=channel1Override, sPlcToNci:=out_stPlcToNci[0]);
ItpSetOverridePercent(fOverridePercent:=channel2Override, sPlcToNci:=out_stPlcToNci[1]);
ItpSetOverridePercent(fOverridePercent:=channel3Override, sPlcToNci:=out_stPlcToNci[2]);

// SetMacro/WaitMacro delle funzioni M: dentro fbMFunc (MacroManager).
// Gruppi e tabelle NC delle sequenze: dentro fbSeq (StateMachine).











udiItpState[0] := ItpGetStateInterpreter(in_stNciToPlc[0]);
udiItpState[1] := ItpGetStateInterpreter(in_stNciToPlc[1]);
udiItpState[2] := ItpGetStateInterpreter(in_stNciToPlc[2]);


fbCloseClampAfterCentering();
ssrActivationDelay();
ssr2ActivationDelay();
waitForMove();
END_ACTION

